(* IEC 61131-3 sources: JingjiangArm/moonboxpro_arm_8.4/Application/Application/任务列表/ExtTask/动作处理/动作处理, 14 files *)

(* ---- KS_ActionBtnDeal.st ---- *)
(*@CES
Name=KS_ActionBtnDeal
Type=FunctionBlock
TypeGuid=6f9dac99-8de1-4efc-8465-68ac443b7d08
Guid=e35c6e03-b7a0-413e-be55-6ff55efa3ce6
HasDeclaration=True
HasImplementation=True
*)
{DECLARATION}
FUNCTION KS_ActionBtnDeal : BOOL
VAR_INPUT
	i_iGrpId								: INT;
	i_pstStEvtReq							: POINTER TO StEvtReq;(*按钮输入操作及边沿触发描述|*)
	i_pbyActionCtlWay						: POINTER TO BYTE;(*动作流程选择
													|0:预启动--空转--张力投入--印刷--空转--停机
													|1:预启动--空转--停机;预启动--张力投入--印刷(速度为0)--停机*)
	i_pxBtnInk								: POINTER TO BOOL;(*空转按钮-包含了预启动响铃状态*)
	i_pxBtnPrint							: POINTER TO BOOL;(*印刷按钮*)
	i_pxBtnTension							: POINTER TO BOOL;(*张力投入按钮*)
	i_pxBtnManuAcc							: POINTER TO BOOL;(*手动加速*)
	i_pxBtnManuDec							: POINTER TO BOOL;(*手动减速*)
	i_pxBtnAutoAccOrDec						: POINTER TO BOOL;(*自动加速减速*)
	i_pxBtnStop								: POINTER TO BOOL;(*停止按钮*)
	i_pxBtnFastStop							: POINTER TO BOOL;(*快速停止按钮|2022.4.9.235931*)
	i_pxBtnEstop							: POINTER TO BOOL;(*急停按钮*)
	i_plrVel_Tar							: POINTER TO LREAL;(*自动加减速目标速度*)

(*2019.09.10.101800|niu.j|*)
	i_xInverterAlarm						: BOOL;(*变频器报警*)
	i_xBrakeFilm							: BOOL;(*断料*)
	(*2022.4.3.165550|*)
	i_xLostPressure							: BOOL;(*气压低报警|不允许开机*)
	i_xPrnRollerLoose_AtLeast1				: BOOL;(*至少一色夹板松报警|不允许开机*)
	i_xNeedEstop_BrakeAlarm					: BOOL;(*制动电阻报警急停|2022.5.11.112758*)
	i_paxCommVel_Sure: POINTER TO ARRAY [1..2,1..3] OF BOOL;
	(*2021.8.27.164750  同步*)
	i_paxNeedRstTrig_AutoAccOrDec:POINTER TO ARRAY [1..3] OF BOOL;(*复位自动加减速按钮沿*)
	i_pxLastFlag_Stop: POINTER TO BOOL;
	i_pxLastFlag_Ink: POINTER TO BOOL;
	i_pxLastFlag_TensionUnFinished:POINTER TO BOOL;(*张力投入未完成标志*)
	i_xFalg_ExhaustEn:BOOL;(*排风启动使能标志|*)
	i_pxFastStopBtnDn:POINTER TO BOOL;(*快停被按下了*)
	i_pxTips_ExhausLimitStart: POINTER TO BOOL;
	i_pbySpecialProcess:POINTER TO BYTE;(*在基础的开机流程上增加了特殊开机方式切换标志|0:按照基础的|
																		 			  |1:北人的*)
	i_ptmHold_PreStart				: POINTER TO TIME; (* 开机预启动持续时间| 2022.5.27.143829*)
	i_tmHold_PreStart_BeiRen		: TIME := T#6s; (* 北人开机预启动持续时间|和响铃时间是分开的| 2022.5.27.143829*)
	i_tmAlarmHold_PreStart			: TIME := t#3s; (* 开机预启动报警持续时间*)
	(*2023.09.21.143646*)
	i_pbyStates						: POINTER TO BYTE;(*状态机@可以在不同厂家独立使用*)
	i_pfbTon						: POINTER TO TON;(*计时器-用于某些流程使用@2023.12.16.151632*)
	i_iCustomerName					: INT;
	i_pxLinkage_IfOf_Ink			: POINTER TO BOOL;
	i_prVel_Tar_HMI					: POINTER TO REAL;(*设定的目标速度值*)
	i_pxTapPosition_Breaking		: POINTER TO BOOL;
	i_pxTapPosition_Printing		: POINTER TO BOOL;
	i_pxTapPosition_UniformInk		: POINTER TO BOOL;
	i_pxAutoAccDec_Hmi				: POINTER TO BOOL;
	i_arVel_CommonlyUsed			: ARRAY [1..3] OF REAL;
	i_xFalg_ExhaustLimitStart		: BOOL;
	i_rVel_Ink						: REAL;
	i_xFlag_Stop					: BOOL;
	i_xFlag_Estop					: BOOL;
	i_xFlag_Ink						: BOOL;
	i_xFlag_Print					: BOOL;
	i_xFlag_InkAccing				: BOOL;
	i_xFlag_Stoping					: BOOL;
	i_xFlag_EStoping				: BOOL;
	i_xFlag_Tension					: BOOL;
	i_xFlag_TensionDone				: BOOL;
	i_xFlag_TensionUnfinished		: BOOL;
	i_xFlag_LinkageAxisAlarm		: BOOL;
	i_rVel_Cur						: REAL;
	i_xFlag_AutoDec					: BOOL;
	i_xFlag_AutoAcc					: BOOL;
	i_xFlag_Accing					: BOOL;
	i_xFlag_Decing					: BOOL;
	i_xMotionEnabled				: BOOL;
	i_pxChangeSts_To_Ink: POINTER TO BOOL;
	i_pxChangeSts_To_Prn: POINTER TO BOOL;
END_VAR
VAR
	iCustomerName: INT;
	iN: INT;
	xInkMove: BOOL;(*空转运动*)
	xNotAllowMachineRun: BOOL;
	xTips_ExhausLimitStart: BOOL;
	xNeedEstopByPrnRollerLoose: BOOL;(*版辊松需要急停*)
	bySpecialProcess:BYTE;(*在基础的开机流程上增加了特殊开机方式切换标志|0:按照基础的|
																		|1:北人的*)
	tmHold_PreStart						: TIME := T#3s; (* 开机预启动持续时间| 2022.5.27.143829*)
	wNotAllowMachineRun:WORD;
	byStates: BYTE;

END_VAR

{IMPLEMENTATION}
KS_ActionBtnDeal:=FALSE;
(*2023.06.24.193214*)
IF i_pbyStates<>0 THEN
	byStates:=i_pbyStates^;
END_IF
IF	i_pstStEvtReq<>0 AND
	i_pbyActionCtlWay<>0 AND
	i_pxBtnInk<>0 AND
	i_pxBtnPrint<>0 AND
	i_pxBtnTension<>0 AND
	i_pxBtnManuAcc<>0 AND
	i_pxBtnManuDec<>0 AND
	i_pxBtnAutoAccOrDec<>0 AND
	i_pxBtnStop<>0 AND
	i_pxBtnFastStop<>0 AND
	i_pxBtnEstop<>0 AND
	i_plrVel_Tar<>0 AND
	i_paxNeedRstTrig_AutoAccOrDec<>0 AND
	i_paxCommVel_Sure<>0 AND
	i_pxFastStopBtnDn<>0 AND
	i_pxChangeSts_To_Ink<>0 AND
	i_pxChangeSts_To_Prn<>0 THEN

	iCustomerName:=i_iCustomerName;(*用户名称*)

	(* 2022.1.11.162754增加牵引联动使能处理*)
	i_pxLinkage_IfOf_Ink^:= TRUE;
	bySpecialProcess:=0;(*默认写0*)
	tmHold_PreStart:=i_tmAlarmHold_PreStart;(*默认赋值*)

	(*2019.10.08.091031|niu.j|按钮复位*)
	i_pxBtnInk^:=FALSE;
	i_pxBtnPrint^:=FALSE;
	i_pxBtnTension^:=FALSE;
	i_pxBtnManuAcc^:=FALSE;
	i_pxBtnManuDec^:=FALSE;
	i_pxBtnAutoAccOrDec^:=FALSE;
	i_pxBtnStop^:=FALSE;
	i_pxBtnFastStop^:=FALSE;
	i_pxBtnEstop^:=FALSE;

	(*2022.4.3.165822  夹板报警|停机 并不允许开机*)
	xNotAllowMachineRun:=FALSE;
	xNeedEstopByPrnRollerLoose:=FALSE;
	wNotAllowMachineRun:= 0;
	IF i_xPrnRollerLoose_AtLeast1 OR
		i_xLostPressure OR
		(NOT i_xFalg_ExhaustEn AND i_xFalg_ExhaustLimitStart) THEN(*排风未启动，限制开机标志使能*)

		IF NOT i_xFlag_Stop AND
			NOT i_xFlag_Estop THEN

			IF i_xPrnRollerLoose_AtLeast1 (*OR(*版辊松就急停*)
				i_xLostPressure*) THEN
				xNeedEstopByPrnRollerLoose:=TRUE;
			END_IF
		ELSE
			IF i_xPrnRollerLoose_AtLeast1 OR(*版辊松*)
				(NOT i_xFalg_ExhaustEn AND i_xFalg_ExhaustLimitStart) OR(*排风限制了不能允许开机*)
				i_xLostPressure THEN(*气压低了也不允许开机@2024.8.17.134512*)
				xNotAllowMachineRun:=TRUE;
				wNotAllowMachineRun.0:= i_xPrnRollerLoose_AtLeast1;(*2022.7.26.102036*)
				wNotAllowMachineRun.1:= (NOT i_xFalg_ExhaustEn AND i_xFalg_ExhaustLimitStart) ;

			END_IF
		END_IF

	END_IF

	(*根据用户名选择开机方式|后期可根据情况将按钮也进行分类2019.9.6.100946*)
	IF i_pbyActionCtlWay<>0 THEN
		CASE iCustomerName OF(*判断用户名称使用不同的开机流程逻辑*)
(*			CUSTOMERNAME_DADONG:
					i_pbyActionCtlWay^:=0;
					(*空转按钮|沿有效*)
					i_pxBtnInk^:=i_pstStEvtReq^.xReqPrestart;
					(*印刷按钮|沿有效*)
					i_pxBtnPrint^:=i_pstStEvtReq^.xReqPrint;
					(*张力投入按钮|沿有效*)
					i_pxBtnTension^:=i_pstStEvtReq^.xReqTension;
					IF i_xFlag_Ink THEN
						(*停止按钮|沿有效*)
						i_pxBtnStop^:=i_pstStEvtReq^.xReqPrestart;
					END_IF
					IF i_xFlag_Print THEN
						(*停止按钮|沿有效*)
						i_pxBtnStop^:=i_pstStEvtReq^.xReqPrint;
					END_IF
					(*无手动加减速*)
					i_pxBtnAutoAccOrDec^:=i_pstStEvtReq^.xReqManuSpdUp OR i_pstStEvtReq^.xReqManuSpdDn;

					IF i_pstStEvtReq^.xReqManuSpdUp THEN(*自动加速了*)
						i_plrVel_Tar^:=i_prVel_Tar_HMI^;
					ELSIF i_pstStEvtReq^.xReqManuSpdDn THEN(*自动减速了|减速到10m/min*)
						i_plrVel_Tar^:= i_rVel_Ink;
					END_IF
					*)
			CUSTOMERNAME_ZHEJIANGOUNUO,(*2023.3.29.114520||增加欧诺*)
			CUSTOMERNAME_SHUNDEDELI,(*2023.10.05.151542*)
			CUSTOMERNAME_BEIREN_NOLOGO,
			CUSTOMERNAME_BEIREN:(*2022.3.24.182915  北人流程*)
					i_pbyActionCtlWay^:=0;
					bySpecialProcess:=1;
					tmHold_PreStart:=i_tmHold_PreStart_BeiRen;
					i_pxBtnFastStop^:=i_pstStEvtReq^.xReqFastStop;(*2022.4.10.000027快停*)
					(*空转按钮|沿有效*)
					(*印刷后空转按钮作为退出印刷状态的按钮*)
					IF i_xFlag_Print THEN
						i_pxBtnStop^:=i_pstStEvtReq^.xReqStop OR i_pstStEvtReq^.xReqInk;
					ELSE
						i_pxBtnStop^:=i_pstStEvtReq^.xReqStop;
						i_pxBtnInk^:=i_pstStEvtReq^.xReqPrestart;
					END_IF

					IF i_pstStEvtReq^.xEvt_FastStop THEN(*快停被按下了*)
						IF i_pxBtnInk^ AND(*开机启动的时候检查下快停按钮输出提示标志*)
							i_xFlag_Stop THEN
							i_pxFastStopBtnDn^:=TRUE;(*快停被按下了*)
							i_pxBtnInk^:=FALSE;(*快停被按下了 就不要开机了*)
						END_IF
					ELSE
						i_pxFastStopBtnDn^:=FALSE;(*快停被按下了*)
					END_IF

					(*印刷按钮|沿有效*)
					i_pxBtnPrint^:=i_pstStEvtReq^.xReqPrint;
					(*张力投入按钮|沿有效*)
					i_pxBtnTension^:=i_pstStEvtReq^.xReqTension;
					(*手动加速|按钮长有效*)
					i_pxBtnManuAcc^:=i_pstStEvtReq^.xEvt_ManuSpdUp;
					(*手动减速|按钮长有效*)
					i_pxBtnManuDec^:=i_pstStEvtReq^.xEvt_ManuSpdDn;
					(*自动加加速|*)
					i_pxBtnAutoAccOrDec^:=i_pstStEvtReq^.xReqPrestart;

					i_plrVel_Tar^:=i_prVel_Tar_HMI^;

					(*2023.09.21.143539 同步*)
					(*2023.3.6.210630 在空转状态下使用空转按键停止到空转速度@我们使用自动减速*)
					IF i_xFlag_Ink AND(*空转状态下*)
						NOT i_xFlag_InkAccing AND(*空转加速完成*)
						NOT (i_xFlag_Stoping OR
						i_xFlag_EStoping) THEN
						IF i_pstStEvtReq^.xReqInk THEN(*空转被按下了*)
							IF i_rVel_Cur>i_rVel_Ink AND
								byStates=0 THEN(*状态为初始值*)
								IF (i_xFlag_AutoAcc OR
									i_xFlag_AutoDec) THEN
									byStates:=2;(*先停止自动加减速再进行自动减速*)
								ELSE(*不在自动加减速中*)
									IF NOT (i_xFlag_Accing OR
										i_xFlag_Decing) THEN(*也不再手动加减速中*)
										byStates:=1;(*自动减速到空转速度*)
									END_IF
								END_IF
							END_IF
						END_IF
					ELSE
						byStates:=0;
					END_IF

					CASE byStates OF
						0:;(*初始值*)
						1:(*自动减速到空转速度*)
							i_pxBtnAutoAccOrDec^:=TRUE;
							i_plrVel_Tar^:=i_rVel_Ink;
							(*忘记了自动加减速按钮按下后几个周期会进入自动加减速状态
							@这里强制等待3个周期认为一定会进入自动加减速状态*)
							byStates:=100;
						2:(*停止自动加减速*)
							i_pxBtnAutoAccOrDec^:=TRUE;
							byStates:=3;(*进入等待一个周期*)
						3:(*等待停止了自动加减速*)
							IF NOT (i_xFlag_Accing OR
								i_xFlag_Decing) THEN(*已经没有加减速了*)
								byStates:=1;(*进入自动减速*)
							END_IF
						100,101:
								byStates:=byStates+1;
								IF byStates=102 THEN
									byStates:=110;(*进入等待步*)
								END_IF
						110:(*等待执行完成@按照逻辑此时应该是会进入自动加减速中*)
							IF i_xFlag_AutoAcc OR
								i_xFlag_AutoDec THEN;
							ELSE(*退出加减速状态的时候复位步*)
								byStates:=0;
							END_IF
					ELSE
						byStates:=0;
					END_CASE

			CUSTOMERNAME_CHENGBAO,
			CUSTOMERNAME_HUAFENG,
			CUSTOMERNAME_SHOUXIN,
			CUSTOMERNAME_RUNXIN,
			CUSTOMERNAME_NBXINDA,
			CUSTOMERNAME_FOSHANCHONGYUAN:
					i_pbyActionCtlWay^:=1;
					IF i_xFlag_Stop THEN
						(*记录下当前的印刷机档位|*)
						i_pxTapPosition_Breaking^:= i_pstStEvtReq^.xEvt_TapPosition_Breaking;
						i_pxTapPosition_Printing^:= i_pstStEvtReq^.xEvt_TapPosition_Printing;
						i_pxTapPosition_UniformInk^:= i_pstStEvtReq^.xEvt_TapPosition_UniformInk;
					END_IF

					IF i_pxTapPosition_Breaking^ THEN(*断料档位*)
						i_pxBtnInk^:=i_pstStEvtReq^.xReqPrestart;(*断料档位只空转*)
					ELSIF i_pxTapPosition_UniformInk^ THEN(*匀墨档位*)
						i_pxBtnInk^:=i_pstStEvtReq^.xReqPrestart;(*匀墨档位-空转+张力投入*)
						IF NOT i_xFlag_Tension THEN
							i_pxBtnTension^:=i_pstStEvtReq^.xReqPrestart;
						END_IF
						i_pxLinkage_IfOf_Ink^:= FALSE;
					ELSIF i_pxTapPosition_Printing^ THEN(*印刷档位*)
						(*印刷档位|在拉料时候有可能会存在牵引电机运动的问题；
						在这里修改启动按钮的时机为拉料完成后|2021.11.3.112006*)

						(*重新优化为先启动电机运动逻辑,再进行拉料@2023.12.16.132911*)
						i_pxBtnPrint^:=i_pstStEvtReq^.xReqPrestart;(*印刷档位-空转+张力投入+印刷0速*)
						IF i_xMotionEnabled THEN
							IF NOT i_xFlag_Tension THEN(*启动拉料*)
								i_pxBtnTension^:=TRUE;
							END_IF
						END_IF
					END_IF

					IF i_pxLastFlag_Stop<>0 THEN
						IF i_xFlag_Tension THEN
							IF (NOT i_xFlag_Estop AND
								i_xFlag_Stop AND
								NOT i_pxLastFlag_Stop^) OR (*非停止到停止*)
								(i_pstStEvtReq^.xReqStop AND
								i_xFlag_Stop) THEN(*停止状态下按下停机按键*)
								i_pxBtnTension^:=TRUE;
								i_pxBtnPrint^:=FALSE;(*和上面逻辑存在状态重叠*)
							END_IF
						END_IF
						i_pxLastFlag_Stop^:=i_xFlag_Stop;

					END_IF

					(*停止按钮|沿有效*)
					i_pxBtnStop^:=i_pstStEvtReq^.xReqStop;
					(*手动加速|按钮长有效*)
					i_pxBtnManuAcc^:=i_pstStEvtReq^.xEvt_ManuSpdUp;
					(*手动减速|按钮长有效*)
					i_pxBtnManuDec^:=i_pstStEvtReq^.xEvt_ManuSpdDn;
					(*自动加加速|*)
					i_pxBtnAutoAccOrDec^:=i_pstStEvtReq^.xReqPrestart;

					i_plrVel_Tar^:=i_prVel_Tar_HMI^;
			CUSTOMERNAME_JIANGYINHUITELI:(*处理江阴汇特力的流程@2023.12.16.133942*)
					i_pbyActionCtlWay^:=1;

					i_pxBtnInk^:=i_pstStEvtReq^.xReqPrestart;(*匀墨档位-空转+张力投入*)
					i_pxBtnPrint^:=i_pstStEvtReq^.xReqPrint;(*印刷按钮*)
					i_pxBtnTension^:=i_pstStEvtReq^.xReqTension;
					(*停止按钮|沿有效*)
					i_pxBtnStop^:=i_pstStEvtReq^.xReqStop;
					(*空转和印刷的时候自动拉张力*)
					IF i_pxLastFlag_Stop<>0 AND i_pbyStates<>0 THEN
						IF (NOT i_xFlag_Estop AND
							NOT i_xFlag_Stop AND
							i_pxLastFlag_Stop^) THEN (*停止到非停止*)
							byStates:=1;(*开机拉张力状态*)
						END_IF
						i_pxLastFlag_Stop^:=i_xFlag_Stop;

						CASE byStates OF
							1:(*开机拉张力*)
								IF NOT i_xFlag_Tension THEN
									i_pxBtnTension^:=TRUE;(*张力投入@等使能都有效了再张力投入*)
								ELSE
									byStates:=2;
								END_IF
							2:(*张力已经启动了*)
								IF i_xFlag_Stop OR
									i_xFlag_EStop THEN
									byStates:=3;
								END_IF
							3:(*取消张力*)
								IF i_xFlag_Tension THEN
									i_pxBtnTension^:=TRUE;
								ELSE(*已经取消了*)
									byStates:=0;
								END_IF
						ELSE
							byStates:=0;
						END_CASE

					END_IF

					(*手动加减速作为自动加减速按钮|按下长达3s就不退出自动加减速-否则退出加减速*)
					IF i_pstStEvtReq^.xEvt_ManuSpdUp AND(*自动加速*)
						i_rVel_Cur<i_prVel_Tar_HMI^ THEN
						i_pxBtnAutoAccOrDec^:=TRUE;
						i_plrVel_Tar^:=i_prVel_Tar_HMI^;
					ELSIF i_pstStEvtReq^.xEvt_ManuSpdDn AND(*自动减速*)
						i_rVel_Cur>0 THEN
						i_pxBtnAutoAccOrDec^:=TRUE;
						i_plrVel_Tar^:=0;
					ELSE
						i_pxBtnAutoAccOrDec^:=FALSE;
						i_plrVel_Tar^:=i_prVel_Tar_HMI^;
					END_IF
					(*自动加减速的时候按下加减速按钮都可以停止@2023.12.17.145038*)
					IF NOT i_pxBtnAutoAccOrDec^ THEN
						IF i_xFlag_AutoAcc OR
							i_xFlag_AutoDec THEN
							i_pxBtnAutoAccOrDec^:=i_pstStEvtReq^.xEvt_ManuSpdUp OR i_pstStEvtReq^.xEvt_ManuSpdDn;
						END_IF
					END_IF

					(*使用计时器计时加减速按钮按下时间决定加速方式@按下3s进入自动加速-否则取消自动加速*)
					IF i_pfbTon<>0 THEN
						IF i_pxBtnAutoAccOrDec^ THEN(*自动加减速按下了*)
							i_pfbTon^(IN:=TRUE,PT:=T#3S);(*启动计时器*)
						ELSE
							IF i_pfbTon^.Q THEN(*时间到了@不处理计时器*)
								IF	NOT(i_xFlag_AutoAcc OR
										i_xFlag_AutoDec) THEN(*退出了自动加减速@复位计时器*)
									i_pfbTon^(IN:=FALSE);(*复位计时器*)
								END_IF
							ELSE(*时间没到|而且按钮取消了,取消自动加减速并复位计时器*)
								IF i_xFlag_AutoAcc OR
									i_xFlag_AutoDec THEN
									IF NOT i_pfbTon^.IN THEN(*用于处理时序@在取消加减速的时候,先复位加减速按钮再置位*)
										i_pxBtnAutoAccOrDec^:=TRUE;
									END_IF
								END_IF
								i_pfbTon^(IN:=FALSE);(*复位计时器*)
							END_IF
						END_IF
					END_IF

			CUSTOMERNAME_ALTMA:
					i_pbyActionCtlWay^:=0;
					(*空转按钮|沿有效*)
					i_pxBtnInk^:=i_pstStEvtReq^.xReqPrestart;
					(*印刷按钮|沿有效*)
					i_pxBtnPrint^:=i_pstStEvtReq^.xReqPrint;
					(*张力投入按钮|沿有效*)
					i_pxBtnTension^:=i_pstStEvtReq^.xReqTension;
					(*停止按钮|沿有效*)
					i_pxBtnStop^:=i_pstStEvtReq^.xReqStop;
					(*手动加速|按钮长有效*)
					i_pxBtnManuAcc^:=i_pstStEvtReq^.xEvt_ManuSpdUp;
					(*手动减速|按钮长有效*)
					i_pxBtnManuDec^:=i_pstStEvtReq^.xEvt_ManuSpdDn;
					(*自动加加速|*)
					i_pxBtnAutoAccOrDec^:=i_pstStEvtReq^.xReqPrestart;
					IF i_xFlag_Ink THEN(*空转时候|空转按键作为自动加速按键*)
						i_pxBtnAutoAccOrDec^:=i_pstStEvtReq^.xReqInk;
					ELSIF i_xFlag_Print THEN(*印刷时候|印刷按键作为自动加速按键*)
						i_pxBtnAutoAccOrDec^:=i_pstStEvtReq^.xReqPrint;
					END_IF

					i_plrVel_Tar^:=i_prVel_Tar_HMI^;

			CUSTOMERNAME_JIANGYINLIDA:(*江阴力达流程修改|2021.12.21.140138*)
					i_pbyActionCtlWay^:=0;
					(*张力投入按钮|沿有效*)
					xInkMove:=i_xFlag_Ink AND
								i_rVel_Cur>0;

					IF i_pxLastFlag_Ink<>0 THEN
						IF  xInkMove AND NOT i_pxLastFlag_Ink^ THEN(*空转以后保证上伺服才能拉料*)
							IF  NOT i_xFlag_Tension THEN
								i_pxBtnTension^:=TRUE;
							END_IF
						END_IF
						i_pxLastFlag_Ink^:=xInkMove;
					END_IF

					IF i_pxLastFlag_Stop<>0 THEN
						IF i_xFlag_Tension THEN
							IF I_xFlag_Stop AND(*停止状态下再按停机|取消张力*)
								i_pstStEvtReq^.xReqStop THEN
								i_pxBtnTension^:=TRUE;
							END_IF
						END_IF
						i_pxLastFlag_Stop^:=i_xFlag_Stop;
					END_IF

					(*空转按钮|沿有效*)
					i_pxBtnInk^:=i_pstStEvtReq^.xReqPrestart;
					(*印刷按钮|沿有效*)
					i_pxBtnPrint^:=i_pstStEvtReq^.xReqPrint;
					(*停止按钮|沿有效*)
					i_pxBtnStop^:=i_pstStEvtReq^.xReqStop;
					(*手动加速|按钮长有效*)
					i_pxBtnManuAcc^:=i_pstStEvtReq^.xEvt_ManuSpdUp;
					(*手动减速|按钮长有效*)
					i_pxBtnManuDec^:=i_pstStEvtReq^.xEvt_ManuSpdDn;
					(*自动加加速|*)
					i_pxBtnAutoAccOrDec^:=i_pstStEvtReq^.xReqPrestart;

					(*张力投入按钮|沿有效*)
					IF NOT i_pxBtnTension^ THEN(* 2021.12.22.144134张力投入按钮*)
						i_pxBtnTension^:=i_pstStEvtReq^.xReqTension;
					END_IF
(* 2021.12.22.145033目标速度赋值*)
					i_plrVel_Tar^:=i_prVel_Tar_HMI^;
			CUSTOMERNAME_JIANGYINHUITONG:(*2022.7.7.102221华丰-流程-类似*)
					i_pbyActionCtlWay^:=0;
					(*空转按钮|沿有效*)
					i_pxBtnInk^:=i_pstStEvtReq^.xReqPrestart;
					(*印刷按钮|沿有效*)
					i_pxBtnPrint^:=i_pstStEvtReq^.xReqPrint;
					(*张力投入按钮|沿有效*)
					i_pxBtnTension^:=i_pstStEvtReq^.xReqTension;
					(*停止按钮|沿有效*)
					i_pxBtnStop^:=i_pstStEvtReq^.xReqStop;
					(*手动加速|按钮长有效*)

					IF i_xFlag_Print THEN(*印刷状态下加速按钮为自动加减速按钮-加减速到目标速度，无手动加速
																，减速为自动减速到空转速度|2022.7.30.093338*)
						i_pxBtnAutoAccOrDec^:= i_pstStEvtReq^.xReqManuSpdUp;(*自动加速*)
						i_plrVel_Tar^:=i_prVel_Tar_HMI^;
						i_pxBtnManuAcc^:=FALSE;(*手动加速无效*)

						IF NOT i_pxBtnAutoAccOrDec^ THEN
							IF i_pstStEvtReq^.xReqManuSpdDn THEN (*手动减速按钮按下-如果速度大于空转速度=自动减速*)
								IF i_rVel_Cur>i_rVel_Ink THEN(*空转速度小于当前速度-自动减速到空转速度*)
									i_pxBtnAutoAccOrDec^:= i_pstStEvtReq^.xReqManuSpdDn;
									i_plrVel_Tar^:=i_rVel_Ink;
								END_IF
							END_IF
						END_IF
					END_IF

					IF i_xFlag_Ink THEN
						IF i_rVel_Cur<i_prVel_Tar_HMI^ THEN(*当前速度小于目标速度-自动加减速生效-手动加减速无效*)
							i_pxBtnAutoAccOrDec^:= i_pstStEvtReq^.xReqManuSpdUp;(*自动加速*)
							i_plrVel_Tar^:=i_prVel_Tar_HMI^;
							i_pxBtnManuAcc^:=FALSE;(*手动加速无效*)
						ELSE
							IF i_xFlag_Ink THEN(*空转有手动加速*)
								i_pxBtnManuAcc^:=i_pstStEvtReq^.xEvt_ManuSpdUp;(*手动加速按钮有效*)
								i_plrVel_Tar^:=i_prVel_Tar_HMI^;
							END_IF
						END_IF

						IF i_pstStEvtReq^.xReqManuSpdDn THEN (*手动减速按钮按下-如果速度大于空转速度=自动减速*)
							IF i_rVel_Cur>i_rVel_Ink THEN(*空转速度小于当前速度-自动减速到空转速度*)
								i_pxBtnAutoAccOrDec^:= i_pstStEvtReq^.xReqManuSpdDn;
								i_plrVel_Tar^:=i_rVel_Ink;
							END_IF
						END_IF
						i_pxBtnManuDec^:=FALSE;(*无手动减速*)
					END_IF
			CUSTOMERNAME_QINHUA:
					i_pbyActionCtlWay^:=1;

					IF i_xFlag_Stop THEN
						(*记录下当前的印刷机档位|*)
						i_pxTapPosition_Breaking^:= i_pstStEvtReq^.xEvt_TapPosition_Breaking;
						i_pxTapPosition_Printing^:= i_pstStEvtReq^.xEvt_TapPosition_Printing;
						i_pxTapPosition_UniformInk^:= i_pstStEvtReq^.xEvt_TapPosition_UniformInk;

						//2026.1.6.160707 | +
						//i_pstStEvtReq^.xReqPrestart := FALSE;
					END_IF

					IF i_pxTapPosition_Breaking^ THEN(*断料档位*)
						i_pxBtnInk^:=i_pstStEvtReq^.xReqPrestart;(*断料档位只空转*)
					ELSIF i_pxTapPosition_UniformInk^ THEN(*匀墨档位*)
						i_pxBtnInk^:=i_pstStEvtReq^.xReqPrestart;(*匀墨档位-空转+张力投入*)
						IF NOT i_xFlag_Tension THEN
							i_pxBtnTension^:=i_pstStEvtReq^.xReqPrestart;
						END_IF
						i_pxLinkage_IfOf_Ink^:= FALSE;
					ELSIF i_pxTapPosition_Printing^ THEN(*印刷档位*)
						(*印刷档位|在拉料时候有可能会存在牵引电机运动的问题；
						在这里修改启动按钮的时机为拉料完成后|2021.11.3.112006*)
(*						i_pxBtnPrint^:=i_pstStEvtReq^.xReqPrestart;(*印刷档位-空转+张力投入+印刷0速*)*)
						IF  NOT i_xFlag_Tension THEN
							i_pxBtnTension^:=i_pstStEvtReq^.xReqPrestart;
						ELSE
							IF  i_xFlag_TensionDone AND (*拉料完成才能进入开机逻辑*)
								i_xFlag_Stop THEN(*停机的时候输出印刷按钮*)
								i_pxBtnPrint^:=TRUE;(*印刷档位-空转+张力投入+印刷0速*)
							END_IF
						END_IF
					END_IF

					IF i_pxLastFlag_Stop<>0 THEN
						IF i_xFlag_Tension THEN
							IF (NOT i_xFlag_Estop AND
								i_xFlag_Stop AND
								NOT i_pxLastFlag_Stop^) OR (*非停止到停止*)
								(i_pstStEvtReq^.xReqStop AND
								i_xFlag_Stop) THEN(*停止状态下按下停机按键*)
								i_pxBtnTension^:=TRUE;
								i_pxBtnPrint^:=FALSE;(*和上面逻辑存在状态重叠*)
							END_IF
						END_IF
						i_pxLastFlag_Stop^:=i_xFlag_Stop;
					END_IF
					(*停止按钮|沿有效*)
					i_pxBtnStop^:=i_pstStEvtReq^.xReqStop;
					(*手动加速|按钮长有效*)
					i_pxBtnManuAcc^:=i_pstStEvtReq^.xEvt_ManuSpdUp;
					(*手动减速|按钮长有效*)
					i_pxBtnManuDec^:=i_pstStEvtReq^.xEvt_ManuSpdDn;
					(*自动加加速|*)
					i_pxBtnAutoAccOrDec^:=i_pstStEvtReq^.xReqPrestart;
					i_plrVel_Tar^:=i_prVel_Tar_HMI^;
			CUSTOMERNAME_CHAOXU:
					i_pbyActionCtlWay^:=1;
					IF i_xFlag_Stop THEN
						(*记录下当前的印刷机档位|*)
						IF i_pxChangeSts_To_Ink^ THEN
							i_pstStEvtReq^.xEvt_TapPosition_UniformInk:= TRUE;
						END_IF

						IF i_pxChangeSts_To_Prn^ THEN
							i_pstStEvtReq^.xEvt_TapPosition_Printing:= TRUE;
						END_IF

						i_pxTapPosition_Breaking^:= i_pstStEvtReq^.xEvt_TapPosition_Breaking;
						i_pxTapPosition_Printing^:= i_pstStEvtReq^.xEvt_TapPosition_Printing;
						i_pxTapPosition_UniformInk^:= i_pstStEvtReq^.xEvt_TapPosition_UniformInk;
					ELSE
						i_pxChangeSts_To_Ink^:= FALSE;
						i_pxChangeSts_To_Prn^:= FALSE;
					END_IF

					IF i_pxTapPosition_Breaking^ THEN(*断料档位*)
						i_pxBtnInk^:=i_pstStEvtReq^.xReqPrestart;(*断料档位只空转*)
					ELSIF i_pxTapPosition_UniformInk^ THEN(*匀墨档位*)
						IF i_xFlag_Tension THEN
							i_pxBtnTension^:= i_pstStEvtReq^.xReqStop;
						END_IF
						IF i_pstStEvtReq^.xReqPrestart THEN
							i_pxChangeSts_To_Prn^:= TRUE;
							i_pxChangeSts_To_Ink^:= FALSE;
							IF NOT i_xFlag_Tension THEN
								i_pxBtnTension^:= i_pstStEvtReq^.xReqPrestart;
							END_IF
						END_IF
						(*
						i_pxBtnInk^:=i_pstStEvtReq^.xReqPrestart;(*匀墨档位-空转+张力投入*)
						IF NOT i_xFlag_Tension THEN
							i_pxBtnTension^:=i_pstStEvtReq^.xReqPrestart;
						END_IF
						i_pxLinkage_IfOf_Ink^:= FALSE;
						*)
					ELSIF i_pxTapPosition_Printing^ THEN(*印刷档位*)
						(*印刷档位|在拉料时候有可能会存在牵引电机运动的问题；
						在这里修改启动按钮的时机为拉料完成后|2021.11.3.112006*)
(*						i_pxBtnPrint^:=i_pstStEvtReq^.xReqPrestart;(*印刷档位-空转+张力投入+印刷0速*)*)
						IF  NOT i_xFlag_Tension THEN
							i_pxBtnTension^:=i_pstStEvtReq^.xReqPrestart;
						ELSE
							IF  i_xFlag_TensionDone AND (*拉料完成才能进入开机逻辑*)
								i_xFlag_Stop THEN(*停机的时候输出印刷按钮*)
								i_pxBtnPrint^:=TRUE;(*印刷档位-空转+张力投入+印刷0速*)
							END_IF
						END_IF
					END_IF

					IF i_pxLastFlag_Stop<>0 THEN
						IF i_xFlag_Tension THEN
							IF (NOT i_xFlag_Estop AND
								i_xFlag_Stop AND
								NOT i_pxLastFlag_Stop^) OR (*非停止到停止*)
								(i_pstStEvtReq^.xReqStop AND
								i_xFlag_Stop) THEN(*停止状态下按下停机按键*)
								//i_pxBtnTension^:=TRUE;
								i_pxChangeSts_To_Ink^:= TRUE;
								i_pxChangeSts_To_Prn^:= FALSE;
								i_pxBtnPrint^:=FALSE;(*和上面逻辑存在状态重叠*)
							END_IF
						END_IF
						i_pxLastFlag_Stop^:=i_xFlag_Stop;
					END_IF

					(*停止按钮|沿有效*)
					i_pxBtnStop^:=i_pstStEvtReq^.xReqStop;
					(*手动加速|按钮长有效*)
					i_pxBtnManuAcc^:=i_pstStEvtReq^.xEvt_ManuSpdUp;
					(*手动减速|按钮长有效*)
					i_pxBtnManuDec^:=i_pstStEvtReq^.xEvt_ManuSpdDn;
					(*自动加加速|*)
					i_pxBtnAutoAccOrDec^:=i_pstStEvtReq^.xReqPrestart;
// 					IF i_xFlag_Print THEN
// 						i_pxBtnAutoAccOrDec^:=i_pstStEvtReq^.xReqPrint;
// 					END_IF
					i_plrVel_Tar^:=i_prVel_Tar_HMI^;
		ELSE
			i_pbyActionCtlWay^:=0;
			(*2023.10.05.152335 将标准开机流程作为默认*)
			(*空转按钮|沿有效*)
			i_pxBtnInk^:=i_pstStEvtReq^.xReqPrestart;
			(*印刷按钮|沿有效*)
			i_pxBtnPrint^:=i_pstStEvtReq^.xReqPrint;
			(*张力投入按钮|沿有效*)
			i_pxBtnTension^:=i_pstStEvtReq^.xReqTension;
			(*停止按钮|沿有效*)
			i_pxBtnStop^:=i_pstStEvtReq^.xReqStop;
			(*手动加速|按钮长有效*)
			i_pxBtnManuAcc^:=i_pstStEvtReq^.xEvt_ManuSpdUp;
			(*手动减速|按钮长有效*)
			i_pxBtnManuDec^:=i_pstStEvtReq^.xEvt_ManuSpdDn;
			(*自动加加速|*)
			i_pxBtnAutoAccOrDec^:=i_pstStEvtReq^.xReqPrestart;

			i_plrVel_Tar^:=i_prVel_Tar_HMI^;

		END_CASE

		IF iCustomerName<> CUSTOMERNAME_BEIREN AND iCustomerName<> CUSTOMERNAME_BEIREN_NOLOGO  AND(*不是北人的流程  清除一些标志*)
			 iCustomerName<> CUSTOMERNAME_ZHEJIANGOUNUO THEN
			i_pxFastStopBtnDn^:=FALSE;
		END_IF

		(*界面自动加减速按钮|2021.7.26.174154*)
		i_pxBtnAutoAccOrDec^:=i_pxBtnAutoAccOrDec^ OR i_pxAutoAccDec_Hmi^;
		i_pxAutoAccDec_Hmi^:=FALSE;

		(*2021.7.17.135538 替换|*)
		FOR iN:=1 TO 3 BY 1 DO
			IF i_paxCommVel_Sure^[i_iGrpId,iN] THEN
(*				i_paxCommVel_Sure^[i_iGrpId,iN]:=FALSE;*)
				i_prVel_Tar_HMI^:=i_arVel_CommonlyUsed[iN];
				IF (NOT i_xFlag_Accing) AND (NOT i_xFlag_Decing) THEN
					IF NOT i_paxNeedRstTrig_AutoAccOrDec^[iN] THEN
						i_paxCommVel_Sure^[i_iGrpId,iN]:=FALSE;
						i_pxBtnAutoAccOrDec^:=TRUE;
					ELSE
						i_paxNeedRstTrig_AutoAccOrDec^[iN]:=FALSE;
						i_pxBtnAutoAccOrDec^:=FALSE;(*2023.12.17.155229@复位处理*)
					END_IF
					i_plrVel_Tar^:=i_prVel_Tar_HMI^;
				ELSE (*自动加速中，停止当前加速启动新加速*)
					IF i_xFlag_AutoAcc  OR i_xFlag_AutoDec THEN
						IF NOT i_pxBtnAutoAccOrDec^ OR i_paxNeedRstTrig_AutoAccOrDec^[iN] THEN(*停止自动加减速*)
							i_pxBtnAutoAccOrDec^:=TRUE;
							i_paxNeedRstTrig_AutoAccOrDec^[iN]:=TRUE;(*还需要再复位一次*)
						ELSIF i_pxBtnAutoAccOrDec^ THEN
							i_paxNeedRstTrig_AutoAccOrDec^[iN]:=TRUE;(*复位沿*)
							i_pxBtnAutoAccOrDec^:=FALSE;(*2023.12.17.155229@复位处理*)
						END_IF
					ELSE
						i_paxCommVel_Sure^[i_iGrpId,iN]:=FALSE;
					END_IF
				END_IF
				EXIT;(*只处理一个有效的*)
			END_IF
		END_FOR

		(*|2022.11.30.093008*)
		(*拉料未完成报警被触发的时候|我们等待拉料完成并再次执行输出印刷按钮启动印刷
		用户不用再按印刷按钮了*)
		IF i_pxLastFlag_TensionUnFinished<>0 THEN
			IF i_xFlag_Tension AND(*处于张力投入中*)
				NOT i_xFlag_Print THEN(*非印刷情况下*)
				IF i_xFlag_TensionUnfinished THEN(*投入未完成|说明按下过印刷*)
					i_pxLastFlag_TensionUnFinished^:=TRUE;
				ELSIF i_pxLastFlag_TensionUnFinished^ AND
					i_xFlag_TensionDone THEN(*张力投入未完成进入到张力投入完成*)
					i_pxBtnPrint^:=TRUE;
					i_pxLastFlag_TensionUnFinished^:=FALSE;
				ELSE(*再按下停止或者急停的时候清除*)
					IF i_pxBtnStop^ OR i_pstStEvtReq^.xEvt_Estop THEN
						i_pxLastFlag_TensionUnFinished^:=FALSE;
					END_IF
				END_IF
			ELSE
				i_pxLastFlag_TensionUnFinished^:=FALSE;
			END_IF
		END_IF
	END_IF

(*
	(*加密处理|2021.12.6.140713*)
	IF g_stEncrytion.Locked THEN
		i_pxBtnPrint^:=FALSE;
	END_IF
*)
	(*急停按钮|沿有效*)
	i_pxBtnEStop^:=	i_pstStEvtReq^.xEvt_Estop OR
						i_xFlag_LinkageAxisAlarm OR
						(i_xInverterAlarm AND (i_xFlag_Print OR i_xFlag_Tension)) OR (* 2021.7.7.171131/ *)
						i_xBrakeFilm (*AND*) OR
(*2022.11.30.092111*)
(*						i_xNeedEstop_BrakeAlarm OR(*2022.5.11.112859*)*)
						xNeedEstopByPrnRollerLoose;(*2022.5.26.165456*)

	(*2022.4.3.170117*)
	IF xNotAllowMachineRun THEN (*不允许开机|*)
		IF i_pxBtnPrint^ OR i_pxBtnInk^ THEN(*2022.5.21.101813|增加排风限制启动提示信息*)
			xTips_ExhausLimitStart:= wNotAllowMachineRun.1;(*TRUE*)(*排风限制启动提示*)
		END_IF
		i_pxBtnInk^:=FALSE;
		i_pxBtnPrint^:=FALSE;
(*		i_pxBtnTension^:=FALSE;*)(*2022.5.21.101039 可以开张力*)
	END_IF

END_IF
(*2022.5.21.102302*)
IF i_pxTips_ExhausLimitStart<>0 THEN
	IF NOT i_pxTips_ExhausLimitStart^ THEN
		IF xTips_ExhausLimitStart THEN(*只置位|*)
			i_pxTips_ExhausLimitStart^:=xTips_ExhausLimitStart;
		END_IF
	ELSE
		IF NOT xNotAllowMachineRun THEN(*机器可以启动了*)
			 i_pxTips_ExhausLimitStart^:=FALSE;
		END_IF
	END_IF
END_IF

(*2022.5.29.001053*)
IF i_pbySpecialProcess<>0 THEN
	i_pbySpecialProcess^:=bySpecialProcess;
END_IF
(*2022.5.29.001053*)
IF i_ptmHold_PreStart<>0 THEN
	i_ptmHold_PreStart^:=tmHold_PreStart;
END_IF

(*2023.06.24.193237*)
IF i_pbyStates<>0 THEN
	i_pbyStates^:=byStates;
END_IF

(* ---- KS_ActionBtnDeal_1.st ---- *)
(*@CES
Name=KS_ActionBtnDeal_1
Type=FunctionBlock
TypeGuid=6f9dac99-8de1-4efc-8465-68ac443b7d08
Guid=29481889-dd1f-4142-86a2-c727a801bd3a
HasDeclaration=True
HasImplementation=True
*)
{DECLARATION}
FUNCTION KS_ActionBtnDeal_1 : BOOL
VAR_INPUT
	i_iGrpId								: INT;
	i_pstStEvtReq							: POINTER TO StEvtReq;(*按钮输入操作及边沿触发描述|*)
	i_pbyActionCtlWay						: POINTER TO BYTE;(*动作流程选择
													|0:预启动--空转--张力投入--印刷--空转--停机
													|1:预启动--空转--停机;预启动--张力投入--印刷(速度为0)--停机*)
	i_pxBtnInk								: POINTER TO BOOL;(*空转按钮-包含了预启动响铃状态*)
	i_pxBtnPrint							: POINTER TO BOOL;(*印刷按钮*)
	i_pxBtnTension							: POINTER TO BOOL;(*张力投入按钮*)
	i_pxBtnManuAcc							: POINTER TO BOOL;(*手动加速*)
	i_pxBtnManuDec							: POINTER TO BOOL;(*手动减速*)
	i_pxBtnAutoAccOrDec						: POINTER TO BOOL;(*自动加速减速*)
	i_pxBtnStop								: POINTER TO BOOL;(*停止按钮*)
	i_pxBtnFastStop							: POINTER TO BOOL;(*快速停止按钮|2022.4.9.235931*)
	i_pxBtnEstop							: POINTER TO BOOL;(*急停按钮*)
	i_plrVel_Tar							: POINTER TO LREAL;(*自动加减速目标速度*)

(*2019.09.10.101800|niu.j|*)
	i_xInverterAlarm						: BOOL;(*变频器报警*)
	i_xBrakeFilm							: BOOL;(*断料*)
	(*2022.4.3.165550|*)
	i_xLostPressure							: BOOL;(*气压低报警|不允许开机*)
	i_xPrnRollerLoose_AtLeast1				: BOOL;(*至少一色夹板松报警|不允许开机*)
	i_xNeedEstop_BrakeAlarm					: BOOL;(*制动电阻报警急停|2022.5.11.112758*)
	i_paxCommVel_Sure: POINTER TO ARRAY [1..2,1..3] OF BOOL;
	(*2021.8.27.164750  同步*)
	i_paxNeedRstTrig_AutoAccOrDec:POINTER TO ARRAY [1..3] OF BOOL;(*复位自动加减速按钮沿*)
	i_pxLastFlag_Stop: POINTER TO BOOL;
	i_pxLastFlag_Ink: POINTER TO BOOL;
	i_pxLastFlag_TensionUnFinished:POINTER TO BOOL;(*张力投入未完成标志*)
	i_xFalg_ExhaustEn:BOOL;(*排风启动使能标志|*)
	i_pxFastStopBtnDn:POINTER TO BOOL;(*快停被按下了*)
	i_pxTips_ExhausLimitStart: POINTER TO BOOL;
	i_pbySpecialProcess:POINTER TO BYTE;(*在基础的开机流程上增加了特殊开机方式切换标志|0:按照基础的|
																		 			  |1:北人的*)
	i_ptmHold_PreStart				: POINTER TO TIME; (* 开机预启动持续时间| 2022.5.27.143829*)
	i_tmHold_PreStart_BeiRen		: TIME := T#6s; (* 北人开机预启动持续时间|和响铃时间是分开的| 2022.5.27.143829*)
	i_tmAlarmHold_PreStart			: TIME := t#3s; (* 开机预启动报警持续时间*)
	(*2023.09.21.143646*)
	i_pbyStates						: POINTER TO BYTE;(*状态机@可以在不同厂家独立使用*)
	i_pfbTon						: POINTER TO TON;(*计时器-用于某些流程使用@2023.12.16.151632*)
	i_iCustomerName					: INT;
	i_pxLinkage_IfOf_Ink			: POINTER TO BOOL;
	i_prVel_Tar_HMI					: POINTER TO REAL;(*设定的目标速度值*)
	i_pxTapPosition_Breaking		: POINTER TO BOOL;
	i_pxTapPosition_Printing		: POINTER TO BOOL;
	i_pxTapPosition_UniformInk		: POINTER TO BOOL;
	i_pxAutoAccDec_Hmi				: POINTER TO BOOL;
	i_arVel_CommonlyUsed			: ARRAY [1..3] OF REAL;
	i_xFalg_ExhaustLimitStart		: BOOL;
	i_rVel_Ink						: REAL;
	i_xFlag_Stop					: BOOL;
	i_xFlag_Estop					: BOOL;
	i_xFlag_Ink						: BOOL;
	i_xFlag_Print					: BOOL;
	i_xFlag_InkAccing				: BOOL;
	i_xFlag_Stoping					: BOOL;
	i_xFlag_EStoping				: BOOL;
	i_xFlag_Tension					: BOOL;
	i_xFlag_TensionDone				: BOOL;
	i_xFlag_TensionUnfinished		: BOOL;
	i_xFlag_LinkageAxisAlarm		: BOOL;
	i_rVel_Cur						: REAL;
	i_xFlag_AutoDec					: BOOL;
	i_xFlag_AutoAcc					: BOOL;
	i_xFlag_Accing					: BOOL;
	i_xFlag_Decing					: BOOL;
	i_xMotionEnabled				: BOOL;
END_VAR
VAR
	iCustomerName: INT;
	iN: INT;
	xInkMove: BOOL;(*空转运动*)
	xNotAllowMachineRun: BOOL;
	xTips_ExhausLimitStart: BOOL;
	xNeedEstopByPrnRollerLoose: BOOL;(*版辊松需要急停*)
	bySpecialProcess:BYTE;(*在基础的开机流程上增加了特殊开机方式切换标志|0:按照基础的|
																		|1:北人的*)
	tmHold_PreStart						: TIME := T#3s; (* 开机预启动持续时间| 2022.5.27.143829*)
	wNotAllowMachineRun:WORD;
	byStates: BYTE;
END_VAR

{IMPLEMENTATION}
KS_ActionBtnDeal:=FALSE;
(*2023.06.24.193214*)
IF i_pbyStates<>0 THEN
	byStates:=i_pbyStates^;
END_IF
IF	i_pstStEvtReq<>0 AND
	i_pbyActionCtlWay<>0 AND
	i_pxBtnInk<>0 AND
	i_pxBtnPrint<>0 AND
	i_pxBtnTension<>0 AND
	i_pxBtnManuAcc<>0 AND
	i_pxBtnManuDec<>0 AND
	i_pxBtnAutoAccOrDec<>0 AND
	i_pxBtnStop<>0 AND
	i_pxBtnFastStop<>0 AND
	i_pxBtnEstop<>0 AND
	i_plrVel_Tar<>0 AND
	i_paxNeedRstTrig_AutoAccOrDec<>0 AND
	i_paxCommVel_Sure<>0 AND
	i_pxFastStopBtnDn<>0 THEN

	iCustomerName:=i_iCustomerName;(*用户名称*)

	(* 2022.1.11.162754增加牵引联动使能处理*)
	i_pxLinkage_IfOf_Ink^:= TRUE;
	bySpecialProcess:=0;(*默认写0*)
	tmHold_PreStart:=i_tmAlarmHold_PreStart;(*默认赋值*)

	(*2019.10.08.091031|niu.j|按钮复位*)
	i_pxBtnInk^:=FALSE;
	i_pxBtnPrint^:=FALSE;
	i_pxBtnTension^:=FALSE;
	i_pxBtnManuAcc^:=FALSE;
	i_pxBtnManuDec^:=FALSE;
	i_pxBtnAutoAccOrDec^:=FALSE;
	i_pxBtnStop^:=FALSE;
	i_pxBtnFastStop^:=FALSE;
	i_pxBtnEstop^:=FALSE;

	(*2022.4.3.165822  夹板报警|停机 并不允许开机*)
	xNotAllowMachineRun:=FALSE;
	xNeedEstopByPrnRollerLoose:=FALSE;
	wNotAllowMachineRun:= 0;
	IF i_xPrnRollerLoose_AtLeast1 OR
		i_xLostPressure OR
		(NOT i_xFalg_ExhaustEn AND i_xFalg_ExhaustLimitStart) THEN(*排风未启动，限制开机标志使能*)

		IF NOT i_xFlag_Stop AND
			NOT i_xFlag_Estop THEN

			IF i_xPrnRollerLoose_AtLeast1 (*OR(*版辊松就急停*)
				i_xLostPressure*) THEN
				xNeedEstopByPrnRollerLoose:=TRUE;
			END_IF
		ELSE
			IF i_xPrnRollerLoose_AtLeast1 OR(*版辊松*)
				(NOT i_xFalg_ExhaustEn AND i_xFalg_ExhaustLimitStart) OR(*排风限制了不能允许开机*)
				i_xLostPressure THEN(*气压低了也不允许开机@2024.8.17.134512*)
				xNotAllowMachineRun:=TRUE;
				wNotAllowMachineRun.0:= i_xPrnRollerLoose_AtLeast1;(*2022.7.26.102036*)
				wNotAllowMachineRun.1:= (NOT i_xFalg_ExhaustEn AND i_xFalg_ExhaustLimitStart) ;

			END_IF
		END_IF

	END_IF

	(*根据用户名选择开机方式|后期可根据情况将按钮也进行分类2019.9.6.100946*)
	IF i_pbyActionCtlWay<>0 THEN
		CASE iCustomerName OF(*判断用户名称使用不同的开机流程逻辑*)
(*			CUSTOMERNAME_DADONG:
					i_pbyActionCtlWay^:=0;
					(*空转按钮|沿有效*)
					i_pxBtnInk^:=i_pstStEvtReq^.xReqPrestart;
					(*印刷按钮|沿有效*)
					i_pxBtnPrint^:=i_pstStEvtReq^.xReqPrint;
					(*张力投入按钮|沿有效*)
					i_pxBtnTension^:=i_pstStEvtReq^.xReqTension;
					IF i_xFlag_Ink THEN
						(*停止按钮|沿有效*)
						i_pxBtnStop^:=i_pstStEvtReq^.xReqPrestart;
					END_IF
					IF i_xFlag_Print THEN
						(*停止按钮|沿有效*)
						i_pxBtnStop^:=i_pstStEvtReq^.xReqPrint;
					END_IF
					(*无手动加减速*)
					i_pxBtnAutoAccOrDec^:=i_pstStEvtReq^.xReqManuSpdUp OR i_pstStEvtReq^.xReqManuSpdDn;

					IF i_pstStEvtReq^.xReqManuSpdUp THEN(*自动加速了*)
						i_plrVel_Tar^:=i_prVel_Tar_HMI^;
					ELSIF i_pstStEvtReq^.xReqManuSpdDn THEN(*自动减速了|减速到10m/min*)
						i_plrVel_Tar^:= i_rVel_Ink;
					END_IF
					*)
			CUSTOMERNAME_ZHEJIANGOUNUO,(*2023.3.29.114520||增加欧诺*)
			CUSTOMERNAME_SHUNDEDELI,(*2023.10.05.151542*)
			CUSTOMERNAME_BEIREN_NOLOGO,
			CUSTOMERNAME_BEIREN:(*2022.3.24.182915  北人流程*)
					i_pbyActionCtlWay^:=0;
					bySpecialProcess:=1;
					tmHold_PreStart:=i_tmHold_PreStart_BeiRen;
					i_pxBtnFastStop^:=i_pstStEvtReq^.xReqFastStop;(*2022.4.10.000027快停*)
					(*空转按钮|沿有效*)
					(*印刷后空转按钮作为退出印刷状态的按钮*)
					IF i_xFlag_Print THEN
						i_pxBtnStop^:=i_pstStEvtReq^.xReqStop OR i_pstStEvtReq^.xReqInk;
					ELSE
						i_pxBtnStop^:=i_pstStEvtReq^.xReqStop;
						i_pxBtnInk^:=i_pstStEvtReq^.xReqPrestart;
					END_IF

					IF i_pstStEvtReq^.xEvt_FastStop THEN(*快停被按下了*)
						IF i_pxBtnInk^ AND(*开机启动的时候检查下快停按钮输出提示标志*)
							i_xFlag_Stop THEN
							i_pxFastStopBtnDn^:=TRUE;(*快停被按下了*)
							i_pxBtnInk^:=FALSE;(*快停被按下了 就不要开机了*)
						END_IF
					ELSE
						i_pxFastStopBtnDn^:=FALSE;(*快停被按下了*)
					END_IF

					(*印刷按钮|沿有效*)
					i_pxBtnPrint^:=i_pstStEvtReq^.xReqPrint;
					(*张力投入按钮|沿有效*)
					i_pxBtnTension^:=i_pstStEvtReq^.xReqTension;
					(*手动加速|按钮长有效*)
					i_pxBtnManuAcc^:=i_pstStEvtReq^.xEvt_ManuSpdUp;
					(*手动减速|按钮长有效*)
					i_pxBtnManuDec^:=i_pstStEvtReq^.xEvt_ManuSpdDn;
					(*自动加加速|*)
					i_pxBtnAutoAccOrDec^:=i_pstStEvtReq^.xReqPrestart;

					i_plrVel_Tar^:=i_prVel_Tar_HMI^;

					(*2023.09.21.143539 同步*)
					(*2023.3.6.210630 在空转状态下使用空转按键停止到空转速度@我们使用自动减速*)
					IF i_xFlag_Ink AND(*空转状态下*)
						NOT i_xFlag_InkAccing AND(*空转加速完成*)
						NOT (i_xFlag_Stoping OR
						i_xFlag_EStoping) THEN
						IF i_pstStEvtReq^.xReqInk THEN(*空转被按下了*)
							IF i_rVel_Cur>i_rVel_Ink AND
								byStates=0 THEN(*状态为初始值*)
								IF (i_xFlag_AutoAcc OR
									i_xFlag_AutoDec) THEN
									byStates:=2;(*先停止自动加减速再进行自动减速*)
								ELSE(*不在自动加减速中*)
									IF NOT (i_xFlag_Accing OR
										i_xFlag_Decing) THEN(*也不再手动加减速中*)
										byStates:=1;(*自动减速到空转速度*)
									END_IF
								END_IF
							END_IF
						END_IF
					ELSE
						byStates:=0;
					END_IF

					CASE byStates OF
						0:;(*初始值*)
						1:(*自动减速到空转速度*)
							i_pxBtnAutoAccOrDec^:=TRUE;
							i_plrVel_Tar^:=i_rVel_Ink;
							(*忘记了自动加减速按钮按下后几个周期会进入自动加减速状态
							@这里强制等待3个周期认为一定会进入自动加减速状态*)
							byStates:=100;
						2:(*停止自动加减速*)
							i_pxBtnAutoAccOrDec^:=TRUE;
							byStates:=3;(*进入等待一个周期*)
						3:(*等待停止了自动加减速*)
							IF NOT (i_xFlag_Accing OR
								i_xFlag_Decing) THEN(*已经没有加减速了*)
								byStates:=1;(*进入自动减速*)
							END_IF
						100,101:
								byStates:=byStates+1;
								IF byStates=102 THEN
									byStates:=110;(*进入等待步*)
								END_IF
						110:(*等待执行完成@按照逻辑此时应该是会进入自动加减速中*)
							IF i_xFlag_AutoAcc OR
								i_xFlag_AutoDec THEN;
							ELSE(*退出加减速状态的时候复位步*)
								byStates:=0;
							END_IF
					ELSE
						byStates:=0;
					END_CASE

			CUSTOMERNAME_CHENGBAO,
			CUSTOMERNAME_HUAFENG,
			CUSTOMERNAME_SHOUXIN,
			CUSTOMERNAME_RUNXIN,
			CUSTOMERNAME_NBXINDA,
			CUSTOMERNAME_FOSHANCHONGYUAN:
					i_pbyActionCtlWay^:=1;
					IF i_xFlag_Stop THEN
						(*记录下当前的印刷机档位|*)
						i_pxTapPosition_Breaking^:= i_pstStEvtReq^.xEvt_TapPosition_Breaking;
						i_pxTapPosition_Printing^:= i_pstStEvtReq^.xEvt_TapPosition_Printing;
						i_pxTapPosition_UniformInk^:= i_pstStEvtReq^.xEvt_TapPosition_UniformInk;
					END_IF

					IF i_pxTapPosition_Breaking^ THEN(*断料档位*)
						i_pxBtnInk^:=i_pstStEvtReq^.xReqPrestart;(*断料档位只空转*)
					ELSIF i_pxTapPosition_UniformInk^ THEN(*匀墨档位*)
						i_pxBtnInk^:=i_pstStEvtReq^.xReqPrestart;(*匀墨档位-空转+张力投入*)
						IF NOT i_xFlag_Tension THEN
							i_pxBtnTension^:=i_pstStEvtReq^.xReqPrestart;
						END_IF
						i_pxLinkage_IfOf_Ink^:= FALSE;
					ELSIF i_pxTapPosition_Printing^ THEN(*印刷档位*)
						(*印刷档位|在拉料时候有可能会存在牵引电机运动的问题；
						在这里修改启动按钮的时机为拉料完成后|2021.11.3.112006*)

						(*重新优化为先启动电机运动逻辑,再进行拉料@2023.12.16.132911*)
						i_pxBtnPrint^:=i_pstStEvtReq^.xReqPrestart;(*印刷档位-空转+张力投入+印刷0速*)
						IF i_xMotionEnabled THEN
							IF NOT i_xFlag_Tension THEN(*启动拉料*)
								i_pxBtnTension^:=TRUE;
							END_IF
						END_IF
					END_IF

					IF i_pxLastFlag_Stop<>0 THEN
						IF i_xFlag_Tension THEN
							IF (NOT i_xFlag_Estop AND
								i_xFlag_Stop AND
								NOT i_pxLastFlag_Stop^) OR (*非停止到停止*)
								(i_pstStEvtReq^.xReqStop AND
								i_xFlag_Stop) THEN(*停止状态下按下停机按键*)
								i_pxBtnTension^:=TRUE;
								i_pxBtnPrint^:=FALSE;(*和上面逻辑存在状态重叠*)
							END_IF
						END_IF
						i_pxLastFlag_Stop^:=i_xFlag_Stop;

					END_IF

					(*停止按钮|沿有效*)
					i_pxBtnStop^:=i_pstStEvtReq^.xReqStop;
					(*手动加速|按钮长有效*)
					i_pxBtnManuAcc^:=i_pstStEvtReq^.xEvt_ManuSpdUp;
					(*手动减速|按钮长有效*)
					i_pxBtnManuDec^:=i_pstStEvtReq^.xEvt_ManuSpdDn;
					(*自动加加速|*)
					i_pxBtnAutoAccOrDec^:=i_pstStEvtReq^.xReqPrestart;

					i_plrVel_Tar^:=i_prVel_Tar_HMI^;
			CUSTOMERNAME_JIANGYINHUITELI:(*处理江阴汇特力的流程@2023.12.16.133942*)
					i_pbyActionCtlWay^:=1;

					i_pxBtnInk^:=i_pstStEvtReq^.xReqPrestart;(*匀墨档位-空转+张力投入*)
					i_pxBtnPrint^:=i_pstStEvtReq^.xReqPrint;(*印刷按钮*)
					i_pxBtnTension^:=i_pstStEvtReq^.xReqTension;
					(*停止按钮|沿有效*)
					i_pxBtnStop^:=i_pstStEvtReq^.xReqStop;
					(*空转和印刷的时候自动拉张力*)
					IF i_pxLastFlag_Stop<>0 AND i_pbyStates<>0 THEN
						IF (NOT i_xFlag_Estop AND
							NOT i_xFlag_Stop AND
							i_pxLastFlag_Stop^) THEN (*停止到非停止*)
							byStates:=1;(*开机拉张力状态*)
						END_IF
						i_pxLastFlag_Stop^:=i_xFlag_Stop;

						CASE byStates OF
							1:(*开机拉张力*)
								IF NOT i_xFlag_Tension THEN
									i_pxBtnTension^:=TRUE;(*张力投入@等使能都有效了再张力投入*)
								ELSE
									byStates:=2;
								END_IF
							2:(*张力已经启动了*)
								IF i_xFlag_Stop OR
									i_xFlag_EStop THEN
									byStates:=3;
								END_IF
							3:(*取消张力*)
								IF i_xFlag_Tension THEN
									i_pxBtnTension^:=TRUE;
								ELSE(*已经取消了*)
									byStates:=0;
								END_IF
						ELSE
							byStates:=0;
						END_CASE

					END_IF

					(*手动加减速作为自动加减速按钮|按下长达3s就不退出自动加减速-否则退出加减速*)
					IF i_pstStEvtReq^.xEvt_ManuSpdUp AND(*自动加速*)
						i_rVel_Cur<i_prVel_Tar_HMI^ THEN
						i_pxBtnAutoAccOrDec^:=TRUE;
						i_plrVel_Tar^:=i_prVel_Tar_HMI^;
					ELSIF i_pstStEvtReq^.xEvt_ManuSpdDn AND(*自动减速*)
						i_rVel_Cur>0 THEN
						i_pxBtnAutoAccOrDec^:=TRUE;
						i_plrVel_Tar^:=0;
					ELSE
						i_pxBtnAutoAccOrDec^:=FALSE;
						i_plrVel_Tar^:=i_prVel_Tar_HMI^;
					END_IF
					(*自动加减速的时候按下加减速按钮都可以停止@2023.12.17.145038*)
					IF NOT i_pxBtnAutoAccOrDec^ THEN
						IF i_xFlag_AutoAcc OR
							i_xFlag_AutoDec THEN
							i_pxBtnAutoAccOrDec^:=i_pstStEvtReq^.xEvt_ManuSpdUp OR i_pstStEvtReq^.xEvt_ManuSpdDn;
						END_IF
					END_IF

					(*使用计时器计时加减速按钮按下时间决定加速方式@按下3s进入自动加速-否则取消自动加速*)
					IF i_pfbTon<>0 THEN
						IF i_pxBtnAutoAccOrDec^ THEN(*自动加减速按下了*)
							i_pfbTon^(IN:=TRUE,PT:=T#3S);(*启动计时器*)
						ELSE
							IF i_pfbTon^.Q THEN(*时间到了@不处理计时器*)
								IF	NOT(i_xFlag_AutoAcc OR
										i_xFlag_AutoDec) THEN(*退出了自动加减速@复位计时器*)
									i_pfbTon^(IN:=FALSE);(*复位计时器*)
								END_IF
							ELSE(*时间没到|而且按钮取消了,取消自动加减速并复位计时器*)
								IF i_xFlag_AutoAcc OR
									i_xFlag_AutoDec THEN
									IF NOT i_pfbTon^.IN THEN(*用于处理时序@在取消加减速的时候,先复位加减速按钮再置位*)
										i_pxBtnAutoAccOrDec^:=TRUE;
									END_IF
								END_IF
								i_pfbTon^(IN:=FALSE);(*复位计时器*)
							END_IF
						END_IF
					END_IF

			CUSTOMERNAME_ALTMA:
					i_pbyActionCtlWay^:=0;
					(*空转按钮|沿有效*)
					i_pxBtnInk^:=i_pstStEvtReq^.xReqPrestart;
					(*印刷按钮|沿有效*)
					i_pxBtnPrint^:=i_pstStEvtReq^.xReqPrint;
					(*张力投入按钮|沿有效*)
					i_pxBtnTension^:=i_pstStEvtReq^.xReqTension;
					(*停止按钮|沿有效*)
					i_pxBtnStop^:=i_pstStEvtReq^.xReqStop;
					(*手动加速|按钮长有效*)
					i_pxBtnManuAcc^:=i_pstStEvtReq^.xEvt_ManuSpdUp;
					(*手动减速|按钮长有效*)
					i_pxBtnManuDec^:=i_pstStEvtReq^.xEvt_ManuSpdDn;
					(*自动加加速|*)
					i_pxBtnAutoAccOrDec^:=i_pstStEvtReq^.xReqPrestart;
					IF i_xFlag_Ink THEN(*空转时候|空转按键作为自动加速按键*)
						i_pxBtnAutoAccOrDec^:=i_pstStEvtReq^.xReqInk;
					ELSIF i_xFlag_Print THEN(*印刷时候|印刷按键作为自动加速按键*)
						i_pxBtnAutoAccOrDec^:=i_pstStEvtReq^.xReqPrint;
					END_IF

					i_plrVel_Tar^:=i_prVel_Tar_HMI^;

			CUSTOMERNAME_JIANGYINLIDA:(*江阴力达流程修改|2021.12.21.140138*)
					i_pbyActionCtlWay^:=0;
					(*张力投入按钮|沿有效*)
					xInkMove:=i_xFlag_Ink AND
								i_rVel_Cur>0;

					IF i_pxLastFlag_Ink<>0 THEN
						IF  xInkMove AND NOT i_pxLastFlag_Ink^ THEN(*空转以后保证上伺服才能拉料*)
							IF  NOT i_xFlag_Tension THEN
								i_pxBtnTension^:=TRUE;
							END_IF
						END_IF
						i_pxLastFlag_Ink^:=xInkMove;
					END_IF

					IF i_pxLastFlag_Stop<>0 THEN
						IF i_xFlag_Tension THEN
							IF I_xFlag_Stop AND(*停止状态下再按停机|取消张力*)
								i_pstStEvtReq^.xReqStop THEN
								i_pxBtnTension^:=TRUE;
							END_IF
						END_IF
						i_pxLastFlag_Stop^:=i_xFlag_Stop;
					END_IF

					(*空转按钮|沿有效*)
					i_pxBtnInk^:=i_pstStEvtReq^.xReqPrestart;
					(*印刷按钮|沿有效*)
					i_pxBtnPrint^:=i_pstStEvtReq^.xReqPrint;
					(*停止按钮|沿有效*)
					i_pxBtnStop^:=i_pstStEvtReq^.xReqStop;
					(*手动加速|按钮长有效*)
					i_pxBtnManuAcc^:=i_pstStEvtReq^.xEvt_ManuSpdUp;
					(*手动减速|按钮长有效*)
					i_pxBtnManuDec^:=i_pstStEvtReq^.xEvt_ManuSpdDn;
					(*自动加加速|*)
					i_pxBtnAutoAccOrDec^:=i_pstStEvtReq^.xReqPrestart;

					(*张力投入按钮|沿有效*)
					IF NOT i_pxBtnTension^ THEN(* 2021.12.22.144134张力投入按钮*)
						i_pxBtnTension^:=i_pstStEvtReq^.xReqTension;
					END_IF
(* 2021.12.22.145033目标速度赋值*)
					i_plrVel_Tar^:=i_prVel_Tar_HMI^;
			CUSTOMERNAME_JIANGYINHUITONG:(*2022.7.7.102221华丰-流程-类似*)
					i_pbyActionCtlWay^:=0;
					(*空转按钮|沿有效*)
					i_pxBtnInk^:=i_pstStEvtReq^.xReqPrestart;
					(*印刷按钮|沿有效*)
					i_pxBtnPrint^:=i_pstStEvtReq^.xReqPrint;
					(*张力投入按钮|沿有效*)
					i_pxBtnTension^:=i_pstStEvtReq^.xReqTension;
					(*停止按钮|沿有效*)
					i_pxBtnStop^:=i_pstStEvtReq^.xReqStop;
					(*手动加速|按钮长有效*)

					IF i_xFlag_Print THEN(*印刷状态下加速按钮为自动加减速按钮-加减速到目标速度，无手动加速
																，减速为自动减速到空转速度|2022.7.30.093338*)
						i_pxBtnAutoAccOrDec^:= i_pstStEvtReq^.xReqManuSpdUp;(*自动加速*)
						i_plrVel_Tar^:=i_prVel_Tar_HMI^;
						i_pxBtnManuAcc^:=FALSE;(*手动加速无效*)

						IF NOT i_pxBtnAutoAccOrDec^ THEN
							IF i_pstStEvtReq^.xReqManuSpdDn THEN (*手动减速按钮按下-如果速度大于空转速度=自动减速*)
								IF i_rVel_Cur>i_rVel_Ink THEN(*空转速度小于当前速度-自动减速到空转速度*)
									i_pxBtnAutoAccOrDec^:= i_pstStEvtReq^.xReqManuSpdDn;
									i_plrVel_Tar^:=i_rVel_Ink;
								END_IF
							END_IF
						END_IF
					END_IF

					IF i_xFlag_Ink THEN
						IF i_rVel_Cur<i_prVel_Tar_HMI^ THEN(*当前速度小于目标速度-自动加减速生效-手动加减速无效*)
							i_pxBtnAutoAccOrDec^:= i_pstStEvtReq^.xReqManuSpdUp;(*自动加速*)
							i_plrVel_Tar^:=i_prVel_Tar_HMI^;
							i_pxBtnManuAcc^:=FALSE;(*手动加速无效*)
						ELSE
							IF i_xFlag_Ink THEN(*空转有手动加速*)
								i_pxBtnManuAcc^:=i_pstStEvtReq^.xEvt_ManuSpdUp;(*手动加速按钮有效*)
								i_plrVel_Tar^:=i_prVel_Tar_HMI^;
							END_IF
						END_IF

						IF i_pstStEvtReq^.xReqManuSpdDn THEN (*手动减速按钮按下-如果速度大于空转速度=自动减速*)
							IF i_rVel_Cur>i_rVel_Ink THEN(*空转速度小于当前速度-自动减速到空转速度*)
								i_pxBtnAutoAccOrDec^:= i_pstStEvtReq^.xReqManuSpdDn;
								i_plrVel_Tar^:=i_rVel_Ink;
							END_IF
						END_IF
						i_pxBtnManuDec^:=FALSE;(*无手动减速*)
					END_IF
			CUSTOMERNAME_QINHUA:
					i_pbyActionCtlWay^:=1;

					IF i_xFlag_Stop THEN
						(*记录下当前的印刷机档位|*)
						i_pxTapPosition_Breaking^:= i_pstStEvtReq^.xEvt_TapPosition_Breaking;
						i_pxTapPosition_Printing^:= i_pstStEvtReq^.xEvt_TapPosition_Printing;
						i_pxTapPosition_UniformInk^:= i_pstStEvtReq^.xEvt_TapPosition_UniformInk;

						//2026.1.6.160707 | +
						//i_pstStEvtReq^.xReqPrestart := FALSE;
					END_IF

					IF i_pxTapPosition_Breaking^ THEN(*断料档位*)
						i_pxBtnInk^:=i_pstStEvtReq^.xReqPrestart;(*断料档位只空转*)
					ELSIF i_pxTapPosition_UniformInk^ THEN(*匀墨档位*)
						i_pxBtnInk^:=i_pstStEvtReq^.xReqPrestart;(*匀墨档位-空转+张力投入*)
						IF NOT i_xFlag_Tension THEN
							i_pxBtnTension^:=i_pstStEvtReq^.xReqPrestart;
						END_IF
						i_pxLinkage_IfOf_Ink^:= FALSE;
					ELSIF i_pxTapPosition_Printing^ THEN(*印刷档位*)
						(*印刷档位|在拉料时候有可能会存在牵引电机运动的问题；
						在这里修改启动按钮的时机为拉料完成后|2021.11.3.112006*)
(*						i_pxBtnPrint^:=i_pstStEvtReq^.xReqPrestart;(*印刷档位-空转+张力投入+印刷0速*)*)
						IF  NOT i_xFlag_Tension THEN
							i_pxBtnTension^:=i_pstStEvtReq^.xReqPrestart;
						ELSE
							IF  i_xFlag_TensionDone AND (*拉料完成才能进入开机逻辑*)
								i_xFlag_Stop THEN(*停机的时候输出印刷按钮*)
								i_pxBtnPrint^:=TRUE;(*印刷档位-空转+张力投入+印刷0速*)
							END_IF
						END_IF
					END_IF

					IF i_pxLastFlag_Stop<>0 THEN
						IF i_xFlag_Tension THEN
							IF (NOT i_xFlag_Estop AND
								i_xFlag_Stop AND
								NOT i_pxLastFlag_Stop^) OR (*非停止到停止*)
								(i_pstStEvtReq^.xReqStop AND
								i_xFlag_Stop) THEN(*停止状态下按下停机按键*)
								i_pxBtnTension^:=TRUE;
								i_pxBtnPrint^:=FALSE;(*和上面逻辑存在状态重叠*)
							END_IF
						END_IF
						i_pxLastFlag_Stop^:=i_xFlag_Stop;
					END_IF
					(*停止按钮|沿有效*)
					i_pxBtnStop^:=i_pstStEvtReq^.xReqStop;
					(*手动加速|按钮长有效*)
					i_pxBtnManuAcc^:=i_pstStEvtReq^.xEvt_ManuSpdUp;
					(*手动减速|按钮长有效*)
					i_pxBtnManuDec^:=i_pstStEvtReq^.xEvt_ManuSpdDn;
					(*自动加加速|*)
					i_pxBtnAutoAccOrDec^:=i_pstStEvtReq^.xReqPrestart;
					i_plrVel_Tar^:=i_prVel_Tar_HMI^;
			CUSTOMERNAME_CHAOXU:
					i_pbyActionCtlWay^:=1;

					IF i_xFlag_Stop THEN
						(*记录下当前的印刷机档位|*)
						i_pxTapPosition_Breaking^:= i_pstStEvtReq^.xEvt_TapPosition_Breaking;
						i_pxTapPosition_Printing^:= i_pstStEvtReq^.xEvt_TapPosition_Printing;
						i_pxTapPosition_UniformInk^:= i_pstStEvtReq^.xEvt_TapPosition_UniformInk;
					END_IF

					IF i_pxTapPosition_Breaking^ THEN(*断料档位*)
						i_pxBtnInk^:=i_pstStEvtReq^.xReqPrestart;(*断料档位只空转*)
					ELSIF i_pxTapPosition_UniformInk^ THEN(*匀墨档位*)
						i_pxBtnInk^:=i_pstStEvtReq^.xReqPrestart;(*匀墨档位-空转+张力投入*)
						IF NOT i_xFlag_Tension THEN
							i_pxBtnTension^:=i_pstStEvtReq^.xReqPrestart;
						END_IF
						i_pxLinkage_IfOf_Ink^:= FALSE;
					ELSIF i_pxTapPosition_Printing^ THEN(*印刷档位*)
						(*印刷档位|在拉料时候有可能会存在牵引电机运动的问题；
						在这里修改启动按钮的时机为拉料完成后|2021.11.3.112006*)
(*						i_pxBtnPrint^:=i_pstStEvtReq^.xReqPrestart;(*印刷档位-空转+张力投入+印刷0速*)*)
						IF  NOT i_xFlag_Tension THEN
							i_pxBtnTension^:=i_pstStEvtReq^.xReqPrestart;
						ELSE
							IF  i_xFlag_TensionDone AND (*拉料完成才能进入开机逻辑*)
								i_xFlag_Stop THEN(*停机的时候输出印刷按钮*)
								i_pxBtnPrint^:=TRUE;(*印刷档位-空转+张力投入+印刷0速*)
							END_IF
						END_IF
					END_IF

					IF i_pxLastFlag_Stop<>0 THEN
						IF i_xFlag_Tension THEN
							IF (NOT i_xFlag_Estop AND
								i_xFlag_Stop AND
								NOT i_pxLastFlag_Stop^) OR (*非停止到停止*)
								(i_pstStEvtReq^.xReqStop AND
								i_xFlag_Stop) THEN(*停止状态下按下停机按键*)
								i_pxBtnTension^:=TRUE;
								i_pxBtnPrint^:=FALSE;(*和上面逻辑存在状态重叠*)
							END_IF
						END_IF
						i_pxLastFlag_Stop^:=i_xFlag_Stop;
					END_IF

					(*停止按钮|沿有效*)
					i_pxBtnStop^:=i_pstStEvtReq^.xReqStop;
					(*手动加速|按钮长有效*)
					i_pxBtnManuAcc^:=i_pstStEvtReq^.xEvt_ManuSpdUp;
					(*手动减速|按钮长有效*)
					i_pxBtnManuDec^:=i_pstStEvtReq^.xEvt_ManuSpdDn;
					(*自动加加速|*)
					i_pxBtnAutoAccOrDec^:=i_pstStEvtReq^.xReqPrestart;
// 					IF i_xFlag_Print THEN
// 						i_pxBtnAutoAccOrDec^:=i_pstStEvtReq^.xReqPrint;
// 					END_IF
					i_plrVel_Tar^:=i_prVel_Tar_HMI^;
		ELSE
			i_pbyActionCtlWay^:=0;
			(*2023.10.05.152335 将标准开机流程作为默认*)
			(*空转按钮|沿有效*)
			i_pxBtnInk^:=i_pstStEvtReq^.xReqPrestart;
			(*印刷按钮|沿有效*)
			i_pxBtnPrint^:=i_pstStEvtReq^.xReqPrint;
			(*张力投入按钮|沿有效*)
			i_pxBtnTension^:=i_pstStEvtReq^.xReqTension;
			(*停止按钮|沿有效*)
			i_pxBtnStop^:=i_pstStEvtReq^.xReqStop;
			(*手动加速|按钮长有效*)
			i_pxBtnManuAcc^:=i_pstStEvtReq^.xEvt_ManuSpdUp;
			(*手动减速|按钮长有效*)
			i_pxBtnManuDec^:=i_pstStEvtReq^.xEvt_ManuSpdDn;
			(*自动加加速|*)
			i_pxBtnAutoAccOrDec^:=i_pstStEvtReq^.xReqPrestart;

			i_plrVel_Tar^:=i_prVel_Tar_HMI^;

		END_CASE

		IF iCustomerName<> CUSTOMERNAME_BEIREN AND iCustomerName<> CUSTOMERNAME_BEIREN_NOLOGO  AND(*不是北人的流程  清除一些标志*)
			 iCustomerName<> CUSTOMERNAME_ZHEJIANGOUNUO THEN
			i_pxFastStopBtnDn^:=FALSE;
		END_IF

		(*界面自动加减速按钮|2021.7.26.174154*)
		i_pxBtnAutoAccOrDec^:=i_pxBtnAutoAccOrDec^ OR i_pxAutoAccDec_Hmi^;
		i_pxAutoAccDec_Hmi^:=FALSE;

		(*2021.7.17.135538 替换|*)
		FOR iN:=1 TO 3 BY 1 DO
			IF i_paxCommVel_Sure^[i_iGrpId,iN] THEN
(*				i_paxCommVel_Sure^[i_iGrpId,iN]:=FALSE;*)
				i_prVel_Tar_HMI^:=i_arVel_CommonlyUsed[iN];
				IF (NOT i_xFlag_Accing) AND (NOT i_xFlag_Decing) THEN
					IF NOT i_paxNeedRstTrig_AutoAccOrDec^[iN] THEN
						i_paxCommVel_Sure^[i_iGrpId,iN]:=FALSE;
						i_pxBtnAutoAccOrDec^:=TRUE;
					ELSE
						i_paxNeedRstTrig_AutoAccOrDec^[iN]:=FALSE;
						i_pxBtnAutoAccOrDec^:=FALSE;(*2023.12.17.155229@复位处理*)
					END_IF
					i_plrVel_Tar^:=i_prVel_Tar_HMI^;
				ELSE (*自动加速中，停止当前加速启动新加速*)
					IF i_xFlag_AutoAcc  OR i_xFlag_AutoDec THEN
						IF NOT i_pxBtnAutoAccOrDec^ OR i_paxNeedRstTrig_AutoAccOrDec^[iN] THEN(*停止自动加减速*)
							i_pxBtnAutoAccOrDec^:=TRUE;
							i_paxNeedRstTrig_AutoAccOrDec^[iN]:=TRUE;(*还需要再复位一次*)
						ELSIF i_pxBtnAutoAccOrDec^ THEN
							i_paxNeedRstTrig_AutoAccOrDec^[iN]:=TRUE;(*复位沿*)
							i_pxBtnAutoAccOrDec^:=FALSE;(*2023.12.17.155229@复位处理*)
						END_IF
					ELSE
						i_paxCommVel_Sure^[i_iGrpId,iN]:=FALSE;
					END_IF
				END_IF
				EXIT;(*只处理一个有效的*)
			END_IF
		END_FOR

		(*|2022.11.30.093008*)
		(*拉料未完成报警被触发的时候|我们等待拉料完成并再次执行输出印刷按钮启动印刷
		用户不用再按印刷按钮了*)
		IF i_pxLastFlag_TensionUnFinished<>0 THEN
			IF i_xFlag_Tension AND(*处于张力投入中*)
				NOT i_xFlag_Print THEN(*非印刷情况下*)
				IF i_xFlag_TensionUnfinished THEN(*投入未完成|说明按下过印刷*)
					i_pxLastFlag_TensionUnFinished^:=TRUE;
				ELSIF i_pxLastFlag_TensionUnFinished^ AND
					i_xFlag_TensionDone THEN(*张力投入未完成进入到张力投入完成*)
					i_pxBtnPrint^:=TRUE;
					i_pxLastFlag_TensionUnFinished^:=FALSE;
				ELSE(*再按下停止或者急停的时候清除*)
					IF i_pxBtnStop^ OR i_pstStEvtReq^.xEvt_Estop THEN
						i_pxLastFlag_TensionUnFinished^:=FALSE;
					END_IF
				END_IF
			ELSE
				i_pxLastFlag_TensionUnFinished^:=FALSE;
			END_IF
		END_IF
	END_IF

(*
	(*加密处理|2021.12.6.140713*)
	IF g_stEncrytion.Locked THEN
		i_pxBtnPrint^:=FALSE;
	END_IF
*)
	(*急停按钮|沿有效*)
	i_pxBtnEStop^:=	i_pstStEvtReq^.xEvt_Estop OR
						i_xFlag_LinkageAxisAlarm OR
						(i_xInverterAlarm AND (i_xFlag_Print OR i_xFlag_Tension)) OR (* 2021.7.7.171131/ *)
						i_xBrakeFilm (*AND*) OR
(*2022.11.30.092111*)
(*						i_xNeedEstop_BrakeAlarm OR(*2022.5.11.112859*)*)
						xNeedEstopByPrnRollerLoose;(*2022.5.26.165456*)

	(*2022.4.3.170117*)
	IF xNotAllowMachineRun THEN (*不允许开机|*)
		IF i_pxBtnPrint^ OR i_pxBtnInk^ THEN(*2022.5.21.101813|增加排风限制启动提示信息*)
			xTips_ExhausLimitStart:= wNotAllowMachineRun.1;(*TRUE*)(*排风限制启动提示*)
		END_IF
		i_pxBtnInk^:=FALSE;
		i_pxBtnPrint^:=FALSE;
(*		i_pxBtnTension^:=FALSE;*)(*2022.5.21.101039 可以开张力*)
	END_IF

END_IF
(*2022.5.21.102302*)
IF i_pxTips_ExhausLimitStart<>0 THEN
	IF NOT i_pxTips_ExhausLimitStart^ THEN
		IF xTips_ExhausLimitStart THEN(*只置位|*)
			i_pxTips_ExhausLimitStart^:=xTips_ExhausLimitStart;
		END_IF
	ELSE
		IF NOT xNotAllowMachineRun THEN(*机器可以启动了*)
			 i_pxTips_ExhausLimitStart^:=FALSE;
		END_IF
	END_IF
END_IF

(*2022.5.29.001053*)
IF i_pbySpecialProcess<>0 THEN
	i_pbySpecialProcess^:=bySpecialProcess;
END_IF
(*2022.5.29.001053*)
IF i_ptmHold_PreStart<>0 THEN
	i_ptmHold_PreStart^:=tmHold_PreStart;
END_IF

(*2023.06.24.193237*)
IF i_pbyStates<>0 THEN
	i_pbyStates^:=byStates;
END_IF

(* ---- KS_ChangeRoller_ValveCTL.st ---- *)
(*@CES
Name=KS_ChangeRoller_ValveCTL
Type=FunctionBlock
TypeGuid=6f9dac99-8de1-4efc-8465-68ac443b7d08
Guid=797ebb41-ab76-4fe9-bfcb-d612c34cdc40
HasDeclaration=True
HasImplementation=True
*)
{DECLARATION}
FUNCTION KS_ChangeRoller_ValveCTL : BOOL(*换版阀控制*)(* 辊子套筒逻辑处理 || 2023.08.01.114908 || bai.zy*)
VAR_INPUT
	i_pastStIOMap_Axis_FE	: POINTER TO ARRAY [1..MAX_UNIT_NUM] OF StIOMap_Axis_FE;(*轴io数据区域|`````````````````````````````````````````````*)
	i_pstStSysParam:POINTER TO StSysParam := 0;(* 整机参数 *)
END_VAR
VAR
	pstStUnitParam_UnSave: POINTER TO StUnitParam_UnSave;(* 色组参数 *)
	pstStIOMap_Axis_FE:POINTER TO StIOMap_Axis_FE;(*轴io数据区域|*)
	iN: INT;
END_VAR
{IMPLEMENTATION}
IF i_pastStIOMap_Axis_FE<>0 AND
	i_pstStSysParam<>0 THEN
	FOR iN:=1 TO i_pstStSysParam^.stStSysParam_Save.iUnitMaxNum BY 1 DO
		pstStUnitParam_UnSave:=ADR(i_pstStSysParam^.astStUnitParam_UnSave[iN]);
		pstStIOMap_Axis_FE:=ADR(i_pastStIOMap_Axis_FE^[iN]);
		(*版辊套筒*)
		pstStIOMap_Axis_FE^.o_xRel_Sleeve_Prn:=FALSE;
		IF pstStUnitParam_UnSave^.rAxisVel_PrnRoller = 0 THEN(*版辊运动了|*)(*版辊不运动时可进行装版 || 2023.08.01.163402 || bai.zy*)
			pstStIOMap_Axis_FE^.o_xRel_Sleeve_Prn:=
						pstStIOMap_Axis_FE^.i_xSleeve_Prn;
		END_IF
		(*网辊套筒*)
		pstStIOMap_Axis_FE^.o_xRel_Sleeve_Net:=FALSE;
		IF pstStUnitParam_UnSave^.rAxisVel_NetRoller = 0 THEN(*网辊运动了|*)(*网辊不运动时可进行装版 || 2023.08.01.163402 || bai.zy*)
			pstStIOMap_Axis_FE^.o_xRel_Sleeve_Net:=
						pstStIOMap_Axis_FE^.i_xSleeve_Net;
		END_IF

	END_FOR
END_IF

(* ---- KS_GetSTime.st ---- *)
(*@CES
Name=KS_GetSTime
Type=FunctionBlock
TypeGuid=6f9dac99-8de1-4efc-8465-68ac443b7d08
Guid=a4f55ea8-3634-425c-a7b6-679c868e638a
HasDeclaration=True
HasImplementation=True
*)
{DECLARATION}
FUNCTION KS_GetSTime : BOOL
(*获取s时间保证加减速前后s时位移一致*)
(*总时间等于速度变化的直线时间+平滑时间*)
VAR_INPUT
	i_byCalcType:BYTE;(*选择平滑时间的方式
								1:按照界面输入的平滑时间和每百米的加速时间设定s曲线;总时间=平滑时间+dv/100*界面时间;平滑时间按照界面设置;
								2:按照比例系数设定平滑时间和每百米的加速时间设定s曲线;总时间=平滑时间+dv/100*界面时间;平滑时间=总时间*系数
								3:按照界面输入加减速时间设定s曲线;总时间=dv/100*界面时间;平滑时间=总时间*系数;
							*)
	i_rSpeed_SCoeff: REAL;(*平滑时间系数@默认2/3*)
	i_iTimeSa_S:INT;(*屏上输入s前时间*)
	i_iTimeEd_S:INT;(*屏上输入s后时间*)
	i_iTime_Acc:INT;(*屏上输入加速时间*)
	i_iTime_Dec:INT;(*屏上输入减速速时间*)
	i_uiMaxVel_UseCalcAcc:UINT;(*计算加速度的速度@100m/min*)
	i_rVel_Cur:REAL;(*当前速度*)
	i_rVel_Tar:REAL;(*目标速度*)
	i_prTimeSa_S:POINTER TO REAL;(*s开始时间*)
	i_prTimeEd_S:POINTER TO REAL;(*s结束时间*)
	i_prDis_Sa:POINTER TO REAL;(*s开始运动的位移*)
	i_prDis_Ed:POINTER TO REAL;(*s结束运动的位移*)
	i_prTime_Total:POINTER TO REAL;(*总时间*)
	i_prTime_SmActual:POINTER TO REAL;(*实际的平滑时间*)
	i_plrTime_Even:POINTER TO LREAL;(*匀加速段的时间@直线加速的时间*)
END_VAR
VAR
	rV0:REAL;
	rVt:REAL;
	rA:REAL;
	rB:REAL;
	rC:REAL;

	byCalcType: BYTE;
	rMaxVel_UseCalcAcc: REAL;
	rTime_AccDec: REAL;(*加减速时间s@界面输入*)
	rTime_S:REAL;(*平滑时间s@以前界面输入是前后,在这里做和处理*)
	rTotalTime: REAL;(*s*)
	rDeltV: REAL;(*m/min*)
	rDeltV_Abs: REAL;(*m/min*)
	rAcceleration_Linear: REAL;(*直线加速度@m/min/s*)
	rAcceleration_Need: REAL;(*实际最大加速度*)
	rTimeSa_S: REAL;(*实际s前时间*)
	rTimeEd_S: REAL;(*实际s后时间*)
	rDis_1: REAL;(*实际s前位移*)
	rDis_2: REAL;(*实际s后位移*)
	rTime_S_Use: REAL;(*实际平滑总时间*)
	rTime_Even:REAL;(*匀加速段的时间*)
END_VAR
{IMPLEMENTATION}
(*计算加速度的速度*)
rMaxVel_UseCalcAcc:=UINT_TO_REAL(i_uiMaxVel_UseCalcAcc);
IF rMaxVel_UseCalcAcc=0 THEN rMaxVel_UseCalcAcc:=100;END_IF
byCalcType:=i_byCalcType;
(*初速度@m/min*)
rV0:=i_rVel_Cur;
(*末速度@m/min*)
rVt:=i_rVel_Tar;
(*速度变化量*)
rDeltV:=rVt-rV0;(*带有方向*)
(*平滑时间*)
rTime_S:=INT_TO_REAL(i_iTimeSa_S+i_iTimeEd_S);

(*加速时间*)
IF rDeltV<0 THEN(*减速*)
	rTime_AccDec:=i_iTime_Dec;
ELSE
	rTime_AccDec:=i_iTime_Acc;
END_IF

IF i_rSpeed_SCoeff =0 THEN
	i_rSpeed_SCoeff:=2.0/3.0;
END_IF

(*rDeltV_Abs:=ABS(rDeltV);(*取正值@计算的是平滑时间*)*)
IF rDeltV<>0 THEN
	IF rTime_AccDec<>0 THEN
		rAcceleration_Linear:=rMaxVel_UseCalcAcc/rTime_AccDec;
	ELSE(*非法值处理*)
		rAcceleration_Linear:=1.5;
	END_IF
	(*需要的总时间@s*)
	rTime_Even:=ABS(rDeltV)/rAcceleration_Linear;(*不会/0*)
	rTotalTime:=rTime_S+rTime_Even;
	IF byCalcType=2 THEN(*总时间=平滑时间+dv/100*界面时间;平滑时间=总时间*系数*)
		rTime_S_Use:=rTotalTime*i_rSpeed_SCoeff;
		rTime_Even:=rTotalTime-rTime_S_Use;
	ELSIF  byCalcType=3 THEN(*总时间=dv/100*界面时间;平滑时间=总时间*系数*)
		rTotalTime:=rTime_Even;
		rTime_S_Use:=rTotalTime*i_rSpeed_SCoeff;
		rTime_Even:=rTotalTime-rTime_S_Use;
	ELSE(*byCalcType=1 默认*)(*总时间=平滑时间+dv/100*界面时间;平滑时间按照界面设置*)
		rTime_S_Use:=rTime_S;
	END_IF
	rAcceleration_Need:=2*rDeltV/(2*rTime_Even+rTime_S_Use);(*不会/0*)

	(*解方程用的A、B、C*)
	rA:=rAcceleration_Need/3.0;(*单位m/min/s*)
	rB:=-rAcceleration_Need*rTime_S_Use/3.0-rV0-rVt;(*单位m/min*)
	rC:=rAcceleration_Need*rTime_S_Use*rTime_S_Use/6.0+rV0*rTime_S_Use;(*m/min*s*)
	(*前后两段的时间*)
	rTimeEd_S:=(-rB-SQRT(rB*rB-4*rA*rC))/2.0/rA;(*单位是s*)
	rTimeSa_S:=rTime_S_Use-rTimeEd_S;

	(*两段时间对应的位移*)
	rDis_1:=rV0*rTimeSa_S+rAcceleration_Need*rTimeSa_S*rTimeSa_S/6.0;(*m/min*s*)
	rDis_1:=rDis_1/60.0;(*m*)
	rDis_2:=rVt*rTimeEd_S-rAcceleration_Need*rTimeEd_S*rTimeEd_S/6.0;
	rDis_2:=rDis_2/60.0;(*m*)
ELSE
	rTimeSa_S:=i_iTimeSa_S;
	rTimeEd_S:=i_iTimeEd_S;
	rTime_Even:=0;
	rDis_1:=0;
	rDis_2:=0;
END_IF
IF i_prTimeSa_S<>0 THEN
	i_prTimeSa_S^:=rTimeSa_S;
END_IF
IF i_prTimeEd_S<>0 THEN
	i_prTimeEd_S^:=rTimeEd_S;
END_IF
IF i_prDis_Sa<>0 THEN
	i_prDis_Sa^:=rDis_1;
END_IF
IF i_prDis_Ed<>0 THEN
	i_prDis_Ed^:=rDis_2;
END_IF
IF i_prTime_Total<>0 THEN
	i_prTime_Total^:=rTotalTime;
END_IF
IF i_prTime_SmActual<>0 THEN
	i_prTime_SmActual^:=rTime_S_Use;
END_IF
IF i_plrTime_Even<>0 THEN
	i_plrTime_Even^:=rTime_Even;
END_IF

(* ---- KS_FB_GetPressDneFlag.st ---- *)
(*@CES
Name=KS_FB_GetPressDneFlag
Type=FunctionBlock
TypeGuid=6f9dac99-8de1-4efc-8465-68ac443b7d08
Guid=5ae664dd-3e73-4120-84fc-3415a767721f
HasDeclaration=True
HasImplementation=True
*)
{DECLARATION}
FUNCTION_BLOCK KS_FB_GetPressDneFlag(*获得压辊实际压刀版辊的标志|放在系流程中*)
VAR_INPUT
	i_xEn: BOOL;
	i_iGrpId: INT;
	i_pstStSysParam: POINTER TO StSysParam;
	i_iGrpAxisNum_Pu: INT; (*印刷色组数*)
	i_aiGrpAxisList: ARRAY [1..MAX_UNIT_NUM] OF INT; (*系的轴列表|已经按照升序排列了*)
	i_pastStIOMap_Main_FE	: POINTER TO ARRAY [1..4] OF StIOMap_Main_FE;(*轴io数据区域|*)
	i_pastStIOMap_Axis_FE	: POINTER TO ARRAY [1..MAX_UNIT_NUM] OF StIOMap_Axis_FE;(*轴io数据区域|`````````````````````````````````````````````*)
	i_paxFlag_PressDne:POINTER TO ARRAY [1..MAX_UNIT_NUM] OF BOOL;(*实际压辊完成标志*)
	i_pxFlag_PressDne_If: POINTER TO BOOL;
	i_pxFlag_PressDne_Of: POINTER TO BOOL;
	i_iAxisId_If: INT;
	i_iAxisId_Of: INT;
	i_iCycleTime_Plc:INT;(*2024.01.22.142644+*)
END_VAR
VAR_OUTPUT
	o_xEn:BOOL;
	o_xRollerStsDn_AtLeast1: BOOL;(*至少一个联动色组合压*)
END_VAR
VAR
	iN: INT;
	iUnitId: INT;
	aiCnt: ARRAY [1..MAX_UNIT_NUM] OF INT;
	iCnt_If: INT;
	iCnt_Of: INT;
	uiTimeMs_RollerPressUpKeep: UINT;
	uiTimeMs_RollerPressUpKeep_If: UINT:= 3000;
	uiTimeMs_RollerPressUpKeep_Of: UINT:= 3000;

	xPressDne: BOOL;

	auiTimeMs_RollerPressUpKeep_In: ARRAY [1..MAX_UNIT_NUM] OF UINT;
	axRel_Press_In: ARRAY [1..MAX_UNIT_NUM] OF BOOL;
	iAxisId_If_In: INT;
	iAxisId_Of_In: INT;
	xRel_Press_If_In: BOOL;
	xRel_Press_Of_In: BOOL;
	axFlag_Linkage_In: ARRAY [1..MAX_UNIT_NUM] OF BOOL;
END_VAR
{IMPLEMENTATION}
o_xEn:=i_xEn;
o_xRollerStsDn_AtLeast1:= FALSE;
IF i_pstStSysParam<>0 AND
	i_pastStIOMap_Main_FE<>0 AND
	i_pastStIOMap_Axis_FE<>0 AND
	i_paxFlag_PressDne<>0 AND
	i_pxFlag_PressDne_If<>0 AND
	i_pxFlag_PressDne_Of<>0 AND
	(i_iGrpId=1 OR i_iGrpId=2) THEN
	(*输入处理一下*)
	iAxisId_If_In:= i_iAxisId_If;
	iAxisId_Of_In:= i_iAxisId_Of;

	IF iAxisId_If_In>0 AND iAxisId_Of_In>0 THEN
		xRel_Press_If_In:= i_pastStIOMap_Main_FE^[iAxisId_If_In].o_xRel_Press_IF;
		xRel_Press_Of_In:= i_pastStIOMap_Main_FE^[iAxisId_Of_In].o_xRel_Press_OF;
	END_IF
	FOR iN:=1 TO MAX_UNIT_NUM BY 1 DO
		auiTimeMs_RollerPressUpKeep_In[iN]:= i_pstStSysParam^.astStUnitParam_Save[iN].uiTimeMs_RollerPressUpKeep;
		axRel_Press_In[iN]:= i_pastStIOMap_Axis_FE^[iN].o_xRel_Press;
		axFlag_Linkage_In[iN]:= i_pstStSysParam^.astStUnitParam_Save[iN].xLinkage;
	END_FOR

	FOR iN:=1 TO MAX_UNIT_NUM BY 1 DO
		IF i_iGrpId=1 THEN(*A系执行在前|我们清除所有输出*)
			i_paxFlag_PressDne^[iN]:=FALSE;
		END_IF
	END_FOR
	i_pxFlag_PressDne_If^:= FALSE;
	i_pxFlag_PressDne_Of^:= FALSE;

	IF i_iCycleTime_Plc<=0 THEN
		i_iCycleTime_Plc:=gc_EXT_TSK_CYCLE_TIME;
	END_IF

	FOR iN:=1 TO i_iGrpAxisNum_Pu BY 1 DO
		iUnitId:=i_aiGrpAxisList[iN];
		IF iUnitId>0 AND iUnitId<=MAX_UNIT_NUM THEN
			uiTimeMs_RollerPressUpKeep:=auiTimeMs_RollerPressUpKeep_In[iUnitId];
			(*最少延时2s判定色组合压完成状态|2020.8.20.203521*)
			(*2022.6.28.145501 调整到3s*)
			IF uiTimeMs_RollerPressUpKeep<=3000 THEN
				uiTimeMs_RollerPressUpKeep:=3000;
			END_IF
			xPressDne:=FALSE;
			IF axRel_Press_In[iUnitId] THEN(*轴合压了*)
				IF aiCnt[iUnitId]*i_iCycleTime_Plc>=uiTimeMs_RollerPressUpKeep THEN
					xPressDne:=TRUE;
				ELSE
					aiCnt[iUnitId]:=aiCnt[iUnitId]+1;
				END_IF
			ELSE
				aiCnt[iUnitId]:=0;
			END_IF

			i_paxFlag_PressDne^[iUnitId]:=xPressDne;
		ELSE;
		END_IF
	END_FOR
	xPressDne:= FALSE;
	IF xRel_Press_If_In THEN
		IF iCnt_If*i_iCycleTime_Plc>=uiTimeMs_RollerPressUpKeep_If THEN
			xPressDne:= TRUE;
		ELSE
			iCnt_If:= iCnt_If+1;
		END_IF
	ELSE
		iCnt_If:= 0;
	END_IF
	i_pxFlag_PressDne_If^:= xPressDne;
	xPressDne:= FALSE;
	IF xRel_Press_Of_In THEN
		IF iCnt_Of*i_iCycleTime_Plc>=uiTimeMs_RollerPressUpKeep_Of THEN
			xPressDne:= TRUE;
		ELSE
			iCnt_Of:= iCnt_Of+1;
		END_IF
	ELSE
		iCnt_Of:= 0;
	END_IF
	i_pxFlag_PressDne_Of^:= xPressDne;

	FOR iN:=1 TO i_iGrpAxisNum_Pu BY 1 DO
		iUnitId:= i_aiGrpAxisList[iN];
		IF axFlag_Linkage_In[iUnitId] AND i_paxFlag_PressDne^[iUnitId] THEN
			IF NOT o_xRollerStsDn_AtLeast1 THEN
				o_xRollerStsDn_AtLeast1:= TRUE;
			END_IF
		END_IF
	END_FOR
END_IF

(* ---- KS_FB_GrpAlarmBellControl.st ---- *)
(*@CES
Name=KS_FB_GrpAlarmBellControl
Type=FunctionBlock
TypeGuid=6f9dac99-8de1-4efc-8465-68ac443b7d08
Guid=91de606a-1433-4ee1-833d-0b9475f7a542
HasDeclaration=True
HasImplementation=True
*)
{DECLARATION}
FUNCTION_BLOCK KS_FB_GrpAlarmBellControl(*报警铃处理功能块|wang.nt|2025.08.12.114029*)
VAR_INPUT
	i_xEn: BOOL;
	i_iGrpId:INT;
	i_iGrpAxisNum_Pu: INT;(*色组轴数|*)
	i_pstStSysParam: POINTER TO StSysParam;
	i_aiGrpAxisList: ARRAY [1..MAX_UNIT_NUM] OF INT;(*轴-站映射表|*)
	i_pastStIOMap_AxisBasic: POINTER TO ARRAY [1..MAX_UNIT_NUM] OF StIOMap_Axis_FE;(*基础io|*)
	i_pastStIOMap_Main: POINTER TO ARRAY [1..MAX_UNIT_NUM] OF StIOMap_Main_FE;(*基础io|*)
	i_pstStEvtReq: POINTER TO StEvtReq;
	i_iAxisId_If: INT;
	i_iAxisId_Of: INT;
	(*乔欣功能增加变量*)
	(*新增加的输入参数--没料时保持响铃，按下任意接料相关按钮则停止响铃|2020.1.10.103514Liu.yt*)
	i_xKeepAlarm_NoMaterial:BOOL;(*有效则一直报警 否则就停止报警！若没有出现过true则按照延迟3s响铃*)
	i_xAlarm_CutDne_Uw:BOOL;(*放料裁切完成后报警一段时间使能标志|5S*)

	(*2020.9.9.115353  针对利佳创增加的报警功能|Liu.yt*)
	i_xAlarm_AccOrDecing:BOOL;
	i_xAlarm_CutFinish_Uw:BOOL;(*接料完成后报警*)
	i_xAlarm_CutFinish_Rw:BOOL;(*接料完成后报警*)
	i_xAlarm_VolDiamAlarm_Uw:BOOL;

	(*2021.4.30.112256 增加放料响铃常输出|*)
	i_xAlarmBell_Uw:BOOL;
	(*2021.6.1.084348 收料报警铃常输出*)
	i_xAlarmBell_Rw:BOOL;
	i_axFlag_AdjValid_V:ARRAY [1..MAX_UNIT_NUM] OF BOOL;(*2025.08.12.150129|纵向自动*)
	i_axThisUnitEna: ARRAY [1..MAX_UNIT_NUM] OF BOOL;(*本色组套色开*)
END_VAR
VAR_OUTPUT
	o_xEno: BOOL;
	o_iErNo: INT;
	o_xPrnRollerLoose_AtLeast1:BOOL;(*至少一色的夹板松了|用于文字提示|2022.4.3.163820*)
	o_xLostPressure:BOOL;(*气压低报警|用于文字提示*)
	o_xbrakeResistanceTempHigh_AtLeast1:BOOL;(*至少一色制动电阻温度高*)
END_VAR
VAR
	iN: INT;
	iAxisId: INT;
	xTmp: BOOL;
	xTmp_UwAlarm: BOOL;
	afbFlag_TON: ARRAY [1..4] OF TON;
	pstStIOMap_AxisBasic: POINTER TO StIOMap_Axis_FE;
	iJ: INT;
	iAxisId_Pu: INT;
	pstStIOMap_Main: POINTER TO StIOMap_Main_FE;

	(*为乔欣没料一直报警以及接料后报警的逻辑添加变量2020.1.10.103803|Liu.yt*)
	xCanAlarm_If: BOOL;
	xFlag_KeepAlarm_NoMaterial: BOOL;
	xFlag_CutDne_Uw: BOOL:=FALSE;
	xCanAlarm_CutDne: BOOL;
	abyLostPressureInCnt: ARRAY [1..MAX_UNIT_NUM] OF BYTE;(*2022.7.24.115721  增加输入防抖*)
	tTimeTmp: TIME;
END_VAR

{IMPLEMENTATION}
o_xEno:= i_xEn;
o_iErNo:= 0;
IF i_xEn THEN
	IF i_iGrpAxisNum_Pu>0 AND
		i_pstStSysParam<>0 AND
		i_pastStIOMap_AxisBasic<>0 AND
		i_pstStEvtReq<>0 THEN

		(*预启动报警|*)
		afbFlag_TON[1](
			IN:= i_pstStSysParam^.astStGrpParam_UnSave[i_iGrpId].xFlag_KeepAlarming,
			PT:= gc_tmAlarmHold_PreStart);

		(*放料卷径报警|*)
		(*2024.8.15.171001+*)
		IF i_pstStSysParam^.stStSysParam_Save.byAlarmHold_VOL_Uw=0 THEN
			i_pstStSysParam^.stStSysParam_Save.byAlarmHold_VOL_Uw:=3;
		END_IF
		tTimeTmp:=DWORD_TO_TIME(BYTE_TO_DWORD(i_pstStSysParam^.stStSysParam_Save.byAlarmHold_VOL_Uw)*1000);

		afbFlag_TON[2](
			IN:= i_pstStSysParam^.astStGrpParam_UnSave[i_iGrpId].xFlag_VolDiamAlarm_Uw,
			PT:= tTimeTmp(*gc_tmAlarmHold_VOL_Uw*));

(*-----------------------------------------------------------------QIAOXIN*)
		(*为乔欣没料一直报警的逻辑添加变量2020.1.10.103555|Liu.yt*)
		IF i_xKeepAlarm_NoMaterial OR
			i_xAlarm_VolDiamAlarm_Uw THEN(*利佳创没料报警标志*)
			xFlag_KeepAlarm_NoMaterial:=TRUE;
		END_IF

		IF xFlag_KeepAlarm_NoMaterial THEN
			xCanAlarm_If:=i_xKeepAlarm_NoMaterial OR i_xAlarm_VolDiamAlarm_Uw;
		ELSE
			xCanAlarm_If:=NOT afbFlag_TON[2].Q;
		END_IF

		(*为乔欣增加的接料后延时5s响铃报警逻辑2020.1.10.103600|Liu.yt*)
		IF i_pstStSysParam^.astStGrpParam_UnSave[i_iGrpId].xFlag_Cut_end_Uw AND i_xAlarm_CutDne_Uw THEN
			xFlag_CutDne_Uw:=TRUE;
		END_IF

		(*2024.8.15.171001+*)
		IF i_pstStSysParam^.stStSysParam_Save.byAlarmHold_CutDne_Uw=0 THEN
			i_pstStSysParam^.stStSysParam_Save.byAlarmHold_CutDne_Uw:=3;
		END_IF
		tTimeTmp:=DWORD_TO_TIME(BYTE_TO_DWORD(i_pstStSysParam^.stStSysParam_Save.byAlarmHold_CutDne_Uw)*1000);

		afbFlag_TON[4](IN:=xFlag_CutDne_Uw,PT:=tTimeTmp(*gc_tmAlarmHold_CutDne_Uw*));(*放料裁切完成*)
		IF afbFlag_TON[4].Q THEN(*时间到了*)
			xFlag_CutDne_Uw:=FALSE;
		END_IF

		xCanAlarm_CutDne:=xFlag_CutDne_Uw;(*启动报警*)

(*-----------------------------------------------------------------QIAOXIN*)

		(*印长报警|*)
		xTmp:= i_pstStSysParam^.astStGrpParam_Save[i_iGrpId].wUwRwAxisProf.1 AND i_pstStSysParam^.astStGrpParam_UnSave[i_iGrpId].axFlag_PrnLen_Alarm[1];
		xTmp:= xTmp OR ((NOT i_pstStSysParam^.astStGrpParam_Save[i_iGrpId].wUwRwAxisProf.1) AND i_pstStSysParam^.astStGrpParam_UnSave[i_iGrpId].axFlag_PrnLen_Alarm[2]);
		xTmp:= xTmp OR i_pstStSysParam^.astStGrpParam_UnSave[i_iGrpId].axFlag_PrnLen_Alarm[3];

		(*2024.8.15.171001+*)
		IF i_pstStSysParam^.stStSysParam_Save.byAlarmHold_PrnLength=0 THEN
			i_pstStSysParam^.stStSysParam_Save.byAlarmHold_PrnLength:=3;
		END_IF
		tTimeTmp:=DWORD_TO_TIME(BYTE_TO_DWORD(i_pstStSysParam^.stStSysParam_Save.byAlarmHold_PrnLength)*1000);

		afbFlag_TON[3](
			IN:= xTmp,
			PT:= tTimeTmp(*gc_tmAlarmHold_PrnLength*));

		IF afbFlag_TON[1].Q AND i_pstStSysParam^.astStGrpParam_UnSave[i_iGrpId].xFlag_KeepAlarming THEN
			i_pstStSysParam^.astStGrpParam_UnSave[i_iGrpId].xFlag_KeepAlarming:= FALSE;
			i_pstStSysParam^.astStGrpParam_UnSave[i_iGrpId].xFlag_PrestartTimeout:=TRUE;
		ELSE
			i_pstStSysParam^.astStGrpParam_UnSave[i_iGrpId].xFlag_PrestartTimeout:=FALSE;
		END_IF

		(*计长报警默认接在收牵处|*)
		xTmp:= (i_pstStSysParam^.astStGrpParam_Save[i_iGrpId].wUwRwAxisProf.1 AND i_pstStSysParam^.astStGrpParam_UnSave[i_iGrpId].axFlag_PrnLen_Alarm[1]);(*A轴印长报警|*)
		xTmp:= xTmp OR ((NOT i_pstStSysParam^.astStGrpParam_Save[i_iGrpId].wUwRwAxisProf.1) AND i_pstStSysParam^.astStGrpParam_UnSave[i_iGrpId].axFlag_PrnLen_Alarm[2]);(*B轴印长报警|*)
		xTmp:= xTmp OR i_pstStSysParam^.astStGrpParam_UnSave[i_iGrpId].axFlag_PrnLen_Alarm[3];(*总印长报警|*)
		IF i_iAxisId_Of>=1 AND i_iAxisId_Of<=MAX_UNIT_NUM THEN
			IF i_pstStSysParam^.astStGrpParam_UnSave[i_iGrpId].xFlag_Print AND
				xTmp AND
				NOT afbFlag_TON[3].Q THEN
				xTmp_UwAlarm:= TRUE;
			ELSE
				xTmp_UwAlarm:= FALSE;
			END_IF
		END_IF

		(*预启动报警或人为按下报警按钮|*)
		IF i_pstStSysParam^.astStGrpParam_UnSave[i_iGrpId].xFlag_KeepAlarming THEN
			xTmp:= TRUE;
		ELSE
			xTmp:= i_pstStEvtReq^.xEvt_AlarmBell;
		END_IF
		xTmp:= xTmp OR xTmp_UwAlarm;

		(*主报警默认接在收牵的位置|*)
		IF i_iAxisId_Of>=1 AND i_iAxisId_Of<=MAX_UNIT_NUM THEN
			pstStIOMap_Main:= ADR(i_pastStIOMap_Main^[i_iAxisId_Of]);
			(*2020.9.9.115605修改下面逻辑屏蔽上面逻辑|Liu.yt*)
			pstStIOMap_Main^.o_xRel_AlarmBell:=xTmp OR
									(i_xAlarm_AccOrDecing OR(*增加了加减速报警2020.9.9.115613*)
									i_xAlarm_CutFinish_Rw) OR(*增加了收料结完料后报警2020.9.9.115618*)
									i_xAlarmBell_Rw;(*2021.6.1.084445 收料报警铃常输出*)

		END_IF

		(*放料报警默认接在放牵处|*)
		IF i_iAxisId_If>=1 AND i_iAxisId_If<=MAX_UNIT_NUM THEN
			pstStIOMap_Main:= ADR(i_pastStIOMap_Main^[i_iAxisId_If]);
			IF (i_pstStSysParam^.astStGrpParam_UnSave[i_iGrpId].xFlag_Print AND
				((i_pstStSysParam^.astStGrpParam_UnSave[i_iGrpId].xFlag_VolDiamAlarm_Uw AND xCanAlarm_If)OR
				i_xAlarm_CutFinish_Uw OR(*放料接料完成报警*)
				xCanAlarm_CutDne)) OR i_xAlarmBell_Uw THEN
				pstStIOMap_Main^.o_xRel_AlarmBell:= TRUE;
			ELSE
				pstStIOMap_Main^.o_xRel_AlarmBell:= FALSE;
			END_IF
		END_IF

		(*2019.01.15.171049|niu.j|套色报警处理*)
		FOR iN:=1 TO i_iGrpAxisNum_Pu BY 1 DO
			iAxisId:= i_aiGrpAxisList[iN];
			pstStIOMap_AxisBasic:= ADR(i_pastStIOMap_AxisBasic^[iAxisId]);
			IF iN<=i_iGrpAxisNum_Pu THEN
				pstStIOMap_AxisBasic^.o_xRel_ArcAlarm_Unit:= FALSE;
				IF i_pstStSysParam^.astStUnitParam_Save[iAxisId].xLinkage AND i_axThisUnitEna[iAxisId] AND i_axFlag_AdjValid_V[iAxisId] THEN
					IF i_pstStSysParam^.astStGrpParam_Save[i_iGrpId].xSwitch_Alarm_Arc THEN
						pstStIOMap_AxisBasic^.o_xRel_ArcAlarm_Unit:= pstStIOMap_AxisBasic^.o_xLamp_Lost
							OR pstStIOMap_AxisBasic^.o_xLamp_Warning;
					ELSE
						;
					END_IF

				END_IF
			ELSE
				pstStIOMap_Main^.o_xRel_ArcAlarm:=FALSE;
				IF i_pstStSysParam^.astStGrpParam_Save[i_iGrpId].xSwitch_Alarm_Arc THEN
					FOR iJ:=1 TO i_iGrpAxisNum_Pu BY 1 DO
						iAxisId_Pu:= i_aiGrpAxisList[iJ];
						pstStIOMap_AxisBasic:= ADR(i_pastStIOMap_AxisBasic^[iAxisId_Pu]);
						IF pstStIOMap_AxisBasic^.o_xRel_ArcAlarm_Unit THEN
							pstStIOMap_Main^.o_xRel_ArcAlarm:= TRUE;
							EXIT;
						ELSE
							;
						END_IF
					END_FOR
				END_IF
			END_IF
		END_FOR

		(*2022.4.3.162946  增加了压力低报警-夹板松报警输出|牵引作为总的夹板松输出*)
		o_xPrnRollerLoose_AtLeast1:=FALSE;
		o_xLostPressure:=FALSE;
		o_xbrakeResistanceTempHigh_AtLeast1:=FALSE;
		FOR iN:=1 TO i_iGrpAxisNum_Pu BY 1 DO
			iAxisId:= i_aiGrpAxisList[iN];
			//pstStAxisParam:= ADR(i_pstStShmGlobalParam^.astStAxisParam[iAxisId]);
			pstStIOMap_AxisBasic:= ADR(i_pastStIOMap_AxisBasic^[iAxisId]);
			(*夹板松报警处理*)
			IF iN<=i_iGrpAxisNum_Pu THEN(*色组轴*)
				pstStIOMap_AxisBasic^.o_xPrnRollerLoose_H:=
									(i_pstStSysParam^.astStUnitParam_Save[iN].xLinkage)AND
									pstStIOMap_AxisBasic^.i_xPrnRollerLoose_H;

				IF NOT o_xPrnRollerLoose_AtLeast1 THEN
					o_xPrnRollerLoose_AtLeast1:=pstStIOMap_AxisBasic^.o_xPrnRollerLoose_H;
				END_IF
			ELSE(*牵引轴*)
				pstStIOMap_AxisBasic^.o_xPrnRollerLoose_H:=o_xPrnRollerLoose_AtLeast1;
			END_IF

			(*气压低报警处理|用于控制响铃*)
			(*2024.8.17.151108 在io获取的地方做了5次防抖*)
			pstStIOMap_AxisBasic^.o_xLostPressure:=pstStIOMap_AxisBasic^.i_xLostPressure;

			IF NOT o_xLostPressure THEN
				o_xLostPressure:=pstStIOMap_AxisBasic^.o_xLostPressure;
			END_IF

			(*ptc过温报警提示*)
			pstStIOMap_AxisBasic^.o_xPtcTempHigh:=pstStIOMap_AxisBasic^.i_xPtcSignal;
			IF NOT o_xbrakeResistanceTempHigh_AtLeast1 THEN
				o_xbrakeResistanceTempHigh_AtLeast1:=pstStIOMap_AxisBasic^.o_xPtcTempHigh;
			END_IF
		END_FOR
	ELSE
		o_iErNo:= -1;
	END_IF
END_IF

(* ---- KS_FB_GrpAxisLinkageCtrl.st ---- *)
(*@CES
Name=KS_FB_GrpAxisLinkageCtrl
Type=FunctionBlock
TypeGuid=6f9dac99-8de1-4efc-8465-68ac443b7d08
Guid=b8bcbe9f-324f-4681-8ae1-7356112ae7c5
HasDeclaration=True
HasImplementation=True
*)
{DECLARATION}
FUNCTION_BLOCK KS_FB_GrpAxisLinkageCtrl
(*2021.10.18.101258  处理界面联动按钮输入|或者从站通讯获得*)
(*2023.10.17.085358 增加至少联动一色标志*)
(*2023.11.27.164625 印刷时候可以切换单联动按钮接口*)
VAR_INPUT
	i_xEn: BOOL;
	i_iGrpId: INT;
	i_iGrpAxisNum_Pu: INT;(*色组轴数|*)
	i_aiGrpAxisList: ARRAY [1..MAX_UNIT_NUM] OF INT;(*轴-站映射表|*)
	i_pstStSysParam: POINTER TO StSysParam;(*整机参数|*)
	i_pastStIOMap_Axis_FE	: POINTER TO ARRAY [1..MAX_UNIT_NUM] OF StIOMap_Axis_FE;(*轴io数据区域|`````````````````````````````````````````````*)
	i_iMaxVel_StsSwitch:INT;(*单联动状态切换的最大速度|2022.7.21.180903*)
	i_xChangLinkageStsWhenPrint:BOOL;(*印刷时候可以切换单联动@2023.11.27.164606*)
END_VAR
VAR_OUTPUT
	o_xEno: BOOL;
	o_iErNo: INT;
	o_xFlag_LinkageAtleast1:BOOL;(*至少联动一色@2023.10.17.085309*)
END_VAR
VAR
	iN: INT;
	pstStUnitParam_Save: POINTER TO StUnitParam_Save;
	pstStUnitParam_UnSave: POINTER TO StUnitParam_UnSave;
	pstStIOMap_Axis_FE: POINTER TO StIOMap_Axis_FE;
	afbR_TRIG: ARRAY [1..MAX_UNIT_NUM] OF R_TRIG;
	axReqLinkage: ARRAY [1..MAX_UNIT_NUM] OF BOOL;
	xTmpResetHomeEnd: BOOL;
	(*2021.10.18.101249  联动按钮界面输入*)
	xLinkageBtn_Hmi: BOOL;
	xLinkageChangeEn: BOOL;(*联动切换使能*)

	iUnitId 	: INT;
(*部分参数需要输入及输出-放这里处理*)
(*输入变量*)
	xAllowLinkageChangeInRunning_In: BOOL;(*在运动过程中允许单联动切换*)
	xFlag_Stop_In: BOOL;
	xFlag_Estop_In: BOOL;
	xFlag_Stoping_In	: BOOL;
	xFlag_FastStoping_In	: BOOL;
	xFlag_EStoping_In		: BOOL;
	xFlag_AllInchRun_In		: BOOL;
	xFlag_Home_In			: BOOL;
	xFlag_PreRegister_In	: BOOL;
	xFlag_PhaseRestore_In	: BOOL;
	xFlag_Print_In			: BOOL;
	rVel_Cur_In				: REAL;
	xUseBtn_Linkage_In			: BOOL;
	axLinkage_IO_In: ARRAY [1..MAX_UNIT_NUM] OF BOOL;(*色组IO联动按钮*)
	axFlag_Alarm_Unit_In: ARRAY [1..MAX_UNIT_NUM] OF BOOL;(*色组报警/离线等标志*)
	xFlag_Alarm_If_In: BOOL;
	xFlag_Alarm_Of_In: BOOL;
	xLinkage_IfOf_Ink_In: BOOL;

(*输出变量*)
	xMoveEnable_Motor_If_Out: BOOL;
	xMoveEnable_Motor_Of_Out: BOOL;
	axLamp_Linkage_IO_Out: ARRAY [1..MAX_UNIT_NUM] OF BOOL;(*色组IO联动指示灯*)
	axMoveEnable_Motor_Out: ARRAY [1..MAX_UNIT_NUM] OF BOOL;(*色组运动使能标志*)
(*输入输出变量*)
	axBtnLinkage_HMI_In_Out: ARRAY [1..MAX_UNIT_NUM] OF BOOL;(*界面联动按钮*)
	axFlag_Linkage_In_Out: ARRAY [1..MAX_UNIT_NUM] OF BOOL;(*色组联动标志*)
	xFlag_Home_end_In_Out: BOOL;
	xFlag_Linkage_If_Out: BOOL;
	xFlag_Linkage_Of_Out: BOOL;

END_VAR
{IMPLEMENTATION}
o_xEno:= i_xEn;
o_iErNo:= 0;
IF i_xEn THEN
	IF i_iGrpAxisNum_Pu>0 AND
		i_pstStSysParam<>0 AND
		i_pastStIOMap_Axis_FE<>0  THEN
		Action_Input();
		(*the parameters are valid|*)
		(*2022.7.8.192719 增加了 单联动切换支持开机逻辑*)
		xLinkageChangeEn:=(xFlag_Stop_In OR xFlag_Estop_In) AND
						(NOT xFlag_Stoping_In) AND
						(NOT xFlag_FastStoping_In) AND(*2022.4.10.000603 快速停止中*)
						(NOT xFlag_EStoping_In) AND
						(NOT xFlag_AllInchRun_In) AND
						(NOT xFlag_Home_In) AND
						(NOT xFlag_PreRegister_In) AND
						(NOT xFlag_PhaseRestore_In);

		IF xAllowLinkageChangeInRunning_In THEN(*支持开机切换单联动*)
			xLinkageChangeEn:=(NOT  xFlag_AllInchRun_In) AND
						(NOT  xFlag_Home_In) AND
						(NOT  xFlag_PreRegister_In) AND
						(NOT  xFlag_PhaseRestore_In)AND
						(*2023.11.27.164834  印刷时候能不能切换增加选择标志*)
						((NOT  xFlag_Print_In AND NOT i_xChangLinkageStsWhenPrint) OR
						i_xChangLinkageStsWhenPrint) AND (*2022.7.21.170040 印刷时候不能切*)
						(rVel_Cur_In<=i_iMaxVel_StsSwitch);(*2022.7.21.180956小于等于切换速度才可以切换*)
		END_IF

(*		IF (i_pstStGrpParam^.xFlag_Stop OR i_pstStGrpParam^.xFlag_Estop) AND
			(NOT i_pstStGrpParam^.xFlag_Stoping) AND
			(NOT i_pstStGrpParam^.xFlag_FastStoping) AND(*2022.4.10.000603 快速停止中*)
			(NOT i_pstStGrpParam^.xFlag_EStoping) AND
			(NOT i_pstStGrpParam^.xFlag_AllInchRun) AND
			(NOT i_pstStGrpParam^.xFlag_Home) AND
			(NOT i_pstStGrpParam^.xFlag_PreRegister) AND
			(NOT i_pstStGrpParam^.xFlag_PhaseRestore) THEN*)
			(*只能在停机的时候转换色组的单联动|*)
		IF  xLinkageChangeEn THEN
			o_xFlag_LinkageAtleast1:=FALSE;(*2023.10.17.085450*)
			FOR iN:=1 TO i_iGrpAxisNum_Pu BY 1 DO
				iUnitId:= i_aiGrpAxisList[iN];(*轴id|*)

				(*2021.10.18.101136 取界面或者从站通讯过来的联动按钮输入|*)
				xLinkageBtn_Hmi:= axBtnLinkage_HMI_In_Out[iUnitId];(*只在按钮控制中起作用*)
				axBtnLinkage_HMI_In_Out[iUnitId]:=FALSE;(*获得之后就清除掉*)
				xTmpResetHomeEnd:= FALSE;

				afbR_TRIG[iN](CLK:=axLinkage_IO_In[iUnitId] OR xLinkageBtn_Hmi, Q=>axReqLinkage[iN]);
				IF xUseBtn_Linkage_In THEN(*非两档开关|*)
					IF axReqLinkage[iN] THEN
						axFlag_Linkage_In_Out[iUnitId]:= NOT axFlag_Linkage_In_Out[iUnitId];
						xTmpResetHomeEnd:= TRUE;
					END_IF
				ELSE
					IF axFlag_Linkage_In_Out[iUnitId]<>axLinkage_IO_In[iUnitId] THEN
						axFlag_Linkage_In_Out[iUnitId]:= axLinkage_IO_In[iUnitId];
						xTmpResetHomeEnd:= TRUE;
					END_IF
				END_IF
				IF xTmpResetHomeEnd AND xFlag_Home_end_In_Out THEN
					xFlag_Home_end_In_Out:= FALSE;
				END_IF
				axLamp_Linkage_IO_Out[iUnitId]:= axFlag_Linkage_In_Out[iUnitId];(*联动指示灯|*)

				axMoveEnable_Motor_Out[iUnitId]:= axFlag_Linkage_In_Out[iUnitId];
				IF xAllowLinkageChangeInRunning_In THEN(*支持开机切换单联动|2022.7.8.193520*)
					IF axFlag_Alarm_Unit_In[iUnitId] THEN(*电机报警了*)
						axMoveEnable_Motor_Out[iUnitId]:=FALSE;
					ELSE
						axMoveEnable_Motor_Out[iUnitId]:=TRUE;(*电机运动使能标志有效|否则根据单联动控制*)
					END_IF
				END_IF

				(*2023.10.17.085232 输出至少联动一色标志*)
				IF axFlag_Linkage_In_Out[iUnitId] THEN
					IF NOT o_xFlag_LinkageAtleast1 THEN
						o_xFlag_LinkageAtleast1:=TRUE;
					END_IF
				END_IF
			END_FOR
		ELSE
			FOR iN:=1 TO MAX_UNIT_NUM BY 1 DO
				iUnitId:= i_aiGrpAxisList[iN];(*轴id|*)
				axBtnLinkage_HMI_In_Out[iUnitId]:=FALSE;(*不能需改的时候单联动状态的时候就清除掉从站发送过来的*)
				afbR_TRIG[iUnitId](CLK:= FALSE);
			END_FOR
		END_IF

		(*牵引|*)
		IF xFlag_Stop_In OR xFlag_Estop_In THEN(*停机或急停都按不联动算|*)
			xFlag_Linkage_If_Out:= FALSE;
			xFlag_Linkage_Of_Out:= FALSE;
		ELSE
			(* 2021.1.14.111720 *)
			IF xFlag_Alarm_If_In THEN
				IF xFlag_Print_In THEN
					xFlag_Linkage_If_Out:= TRUE;
				END_IF
			ELSE
				(* 2022.1.11.162926增加牵引空转使能*)
				IF xLinkage_IfOf_Ink_In THEN
					xFlag_Linkage_If_Out:= xLinkage_IfOf_Ink_In;
					(*pstStAxisParam^.xLinkage:= TRUE;*)
				END_IF
			END_IF
			(* 2021.1.14.111720 *)
			IF xFlag_Alarm_Of_In THEN
				IF xFlag_Print_In THEN
					xFlag_Linkage_Of_Out:= TRUE;
				END_IF
			ELSE
				(* 2022.1.11.162926增加牵引空转使能*)
				IF xLinkage_IfOf_Ink_In THEN
					xFlag_Linkage_Of_Out:= xLinkage_IfOf_Ink_In;
					(*pstStAxisParam^.xLinkage:= TRUE;*)
				END_IF
			END_IF
		END_IF
		xMoveEnable_Motor_If_Out:=xFlag_Linkage_If_Out;(*少了这行代码*)
		xMoveEnable_Motor_Of_Out:=xFlag_Linkage_Of_Out;(*少了这行代码*)
		Action_Output();

	ELSE
		o_iErNo:= -1;
		o_xFlag_LinkageAtleast1:=FALSE;(*2023.10.17.085450*)
	END_IF
ELSE
	o_xFlag_LinkageAtleast1:=FALSE;(*2023.10.17.085450*)
END_IF
